(* Collect hmi signals *)
stgGr05HMI.stPLCTOHMI.bHomeCompleted := bgGr05HomeCompleted;
stgGr05HMI.stPLCTOHMI.wBtnStartStatus.0 := bgGr05StartProcess;
stgGr05HMI.stPLCTOHMI.wBtnStopStatus.0 := NOT bgGr05StartProcess;
stgGr05HMI.stPLCTOHMI.wBtnStepProcStatus := 0;
stgGr05HMI.stPLCTOHMI.wAxisClampStatus.0 := NOT binGr05AxisClamp1LimitMin;
stgGr05HMI.stPLCTOHMI.wAxisClampStatus.1 := NOT binGr05AxisClamp1LimitMax;
stgGr05HMI.stPLCTOHMI.wSlideStatus.0 := binGr05SlideTop;
stgGr05HMI.stPLCTOHMI.wSlideStatus.1 := binGr05SlideBottom;
stgGr05HMI.stPLCTOHMI.wRemovalBandStatus.0 := NOT binGr05RemovalBandInMinus;
stgGr05HMI.stPLCTOHMI.wRemovalBandStatus.1 := NOT binGr05RemovalBandInPlus;
stgGr05HMI.stPLCTOHMI.arwClampStatus[1].0 := arbinGr05ClampOpened[1];
stgGr05HMI.stPLCTOHMI.arwClampStatus[1].1 := arbinGr05ClampClosed[1];
stgGr05HMI.stPLCTOHMI.arwClampStatus[2].0 := arbinGr05ClampOpened[2];
stgGr05HMI.stPLCTOHMI.arwClampStatus[2].1 := arbinGr05ClampClosed[2];
stgGr05HMI.stPLCTOHMI.arwCylinderPosStatus[1].0 := arbinGr05CylinderPosOpened[1];
stgGr05HMI.stPLCTOHMI.arwCylinderPosStatus[1].1 := arbinGr05CylinderPosClosed[1];
stgGr05HMI.stPLCTOHMI.arwCylinderPosStatus[2].0 := arbinGr05CylinderPosOpened[2];
stgGr05HMI.stPLCTOHMI.arwCylinderPosStatus[2].1 := arbinGr05CylinderPosClosed[2];
stgGr05HMI.stPLCTOHMI.arwCylinderPosStatus[3].0 := arbinGr05CylinderPosOpened[3];
stgGr05HMI.stPLCTOHMI.arwCylinderPosStatus[3].1 := arbinGr05CylinderPosClosed[3];
stgGr05HMI.stPLCTOHMI.unSawingStep := Gr05Auto.fbProcedure.unProcessCounter;
END_ACTION

END_PROGRAM

// ---- POUs/Tc2 Objects/MachineEquipment/F_AxisClamp2Pos.TcPOU
FUNCTION F_AxisClamp2Pos : LREAL
(*

The function  used to generate position position dependent of diameter and angle.

Constructor: 		Patryk Panylo
Company:		E. Riexinger GmbH
Date:			01.04.2015
Version:			1.00

Date:			Revision:		Who:				Comment
dd.mm.yyyy		x.xx			Initials			comment

*)
VAR_INPUT
	(* Input variables / Eingang Variablen *)
	bEnable							:BOOL;						(* Function block enable *)
	lrActClamp2Pos					:LREAL;
	lrAngle							:LREAL;
	lrRadius							:LREAL;
	lrPipeClampWidth					:LREAL;
	lrSawbandGuideWidth				:LREAL;
END_VAR
VAR
	lrOffset : LREAL;
END_VAR

IF NOT bEnable
THEN
	F_AxisClamp2Pos := lrActClamp2Pos;
	RETURN;
END_IF

lrAngle := LIMIT(-45, lrAngle, 45);



F_AxisClamp2Pos := (TAN(ABS(lrAngle)) * (lrRadius + lrPipeClampWidth))
				     + (lrSawbandGuideWidth / 2 / COS(ABS(lrAngle)))
				     - (lrSawbandGuideWidth / 2);

END_FUNCTION

// ---- POUs/Tc2 Objects/Basics/FB_CheckArrayBounds.TcPOU
FUNCTION_BLOCK FB_CheckArrayBounds
VAR_INPUT
	diArrayIndex: DINT;
	diLowerBound: DINT;
	diUpperBound: DINT;
END_VAR
VAR_OUTPUT
	sLogMessage: STRING;
	diReturnBound: DINT;
END_VAR
VAR
	bErrorUpper: BOOL;
	bErrorLower: BOOL;
	fbRTrig_MessageOutputLower: R_TRIG;
	fbRTrig_MessageOutputUpper: R_TRIG;
END_VAR

(*++++++++++ Checkbounds ++++++++++*)
(*If somehow it happens that a value of any of the used arrays that does not exist is being accessed,
the value is either set to the highest declared value (if a value higher than the highest declared value is being accessed) 
or it is set to the lowest declared value (if a value lower than the lowest declared value is being accessed)  *)

IF diArrayIndex< diLowerBound THEN
	diReturnBound:= diLowerBound;
	bErrorLower:= TRUE;

	sLogMessage:= 'CheckBounds: Array index too LOW! Lower Bound: ';			(*Message is put together*)
	sLogMessage:=CONCAT(sLogMessage,DINT_TO_STRING(diLowerBound));
	sLogMessage:=CONCAT(sLogMessage,' Index being accessed: ');
	sLogMessage:=CONCAT(sLogMessage,DINT_TO_STRING(diArrayIndex));

ELSIF diArrayIndex> diUpperBound THEN
	diReturnBound:= diUpperBound;
	bErrorUpper:= TRUE;

	sLogMessage:= 'CheckBounds: Array index too HIGH! Upper Bound: ';			(*Message is put together*)
	sLogMessage:=CONCAT(sLogMessage,DINT_TO_STRING(diUpperBound));
	sLogMessage:=CONCAT(sLogMessage,' Index being accessed: ');
	sLogMessage:=CONCAT(sLogMessage,DINT_TO_STRING(diArrayIndex));

ELSIF NOT (diArrayIndex< diLowerBound) AND
	NOT (diArrayIndex> diUpperBound) THEN
		diReturnBound:= diArrayIndex;
		bErrorUpper:= FALSE;
		bErrorLower:= FALSE;
END_IF

(*++++++++++ ADSLOGDINT ++++++++++*)
(*If somehow it happens that a value of any of the used arrays that does not exist is being accessed,
the Error is written into the Logger Box of the TC System Manager  *)

fbRTrig_MessageOutputLower( CLK:= bErrorLower, Q=> );
fbRTrig_MessageOutputUpper( CLK:= bErrorUpper, Q=> );

IF fbRTrig_MessageOutputLower.Q OR fbRTrig_MessageOutputUpper.Q THEN
	ADSLOGDINT( ADSLOG_MSGTYPE_ERROR OR ADSLOG_MSGTYPE_LOG,sLogMessage,0);	(*Message is written into Event Log*)
END_IF

END_FUNCTION_BLOCK

// ---- POUs/Tc2 Objects/Basics/CheckBounds.TcPOU
FUNCTION CheckBounds : DINT
VAR_INPUT
	index: DINT;
	lower: DINT;
	upper: DINT;
END_VAR
VAR_EXTERNAL
	fbCheckArrayBounds: FB_CheckArrayBounds;
END_VAR

(*This function checks if an index out of range an array is being accessed *)

fbCheckArrayBounds(
	diArrayIndex			:= index,
	diLowerBound		:= lower,
	diUpperBound		:= upper,
	sLogMessage		=> ,
	diReturnBound		=> CheckBounds);

END_FUNCTION

// ---- POUs/Tc2 Objects/Basics/FB_CheckDivRealInfo.TcPOU
FUNCTION_BLOCK FB_CheckDivRealInfo
VAR_INPUT
	rDivisor: REAL;
END_VAR
VAR_OUTPUT
	rReturnDivReal: REAL;
	sLogMessage: STRING;
END_VAR
VAR
	bDivisorError: BOOL;
	fbRTrig_MessageOutputDiv: R_TRIG;
END_VAR

IF rDivisor= 0 THEN
	bDivisorError:= TRUE;
	rReturnDivReal:= 1;
ELSE
	rReturnDivReal:= rDivisor;
	bDivisorError:= FALSE;
END_IF

(*++++++++++ ADSLOGDINT ++++++++++*)
(*If somewhere a division by 0 is performed, an Error is written into the Logger Box of the TC System Manager  *)

fbRTrig_MessageOutputDiv( CLK:= bDivisorError, Q=> );

IF fbRTrig_MessageOutputDiv.Q THEN
	sLogMessage:= 'CheckDivReal Error: Division by Zero! Divisor set from 0 to 1. ';					(*Message*)

	ADSLOGDINT( ADSLOG_MSGTYPE_ERROR OR ADSLOG_MSGTYPE_LOG,sLogMessage,0);	(*Message is written into Event Log*)
END_IF

END_FUNCTION_BLOCK

// ---- POUs/Tc2 Objects/Basics/CheckDivReal.TcPOU
FUNCTION CheckDivReal : REAL
VAR_INPUT
	divisor: REAL;
END_VAR
VAR_EXTERNAL
	fbCheckDivRealInfo: FB_CheckDivRealInfo;
END_VAR

(*This function checks if a division by zero is performed*)

fbCheckDivRealInfo(
	rDivisor			:= divisor,
	sLogMessage	=> ,
	rReturnDivReal 	=> CheckDivReal);

END_FUNCTION

// ---- POUs/FAST.TcPOU
PROGRAM FAST
VAR
	(* Enummerations *)

	(* Variables *)

	(* References *)

	(* Interfaces *)

	(* Instances *)

END_VAR


;

END_PROGRAM

// ---- POUs/Tc2 Objects/Automation/Axis/Beckhoff/FB_AxisMcBeckhoff.TcPOU
FUNCTION_BLOCK FB_AxisMcBeckhoff
(*

The function block used to control axis welding.

Constructor: 		Patryk Panylo
Company:		E. Riexinger GmbH
Date:			28.04.2015
Version:			1.00

Date:			Revision:		Who:				Comment
dd.mm.yyyy		x.xx			Initials			comment

*)
VAR_INPUT
	(* Input variables / Eingang Variablen *)
	bEnable						:BOOL;						(* Axis present *)
	etMachineMode				:ET_MachineMode;			(* Machine mode *)
	etMachineState				:ET_MachineState;			(* Machine state *)
	bNoEStop					:BOOL;						(* No ermergency Stop / Keine Notaus *)
	bPowerSupplyOn				:BOOL;						(* Power supply on / Leitung eingeschaltet *)
	bLightCurtainOK				:BOOL;						(* Light curtain ok / Freigabe Lichtschranke i.o *)
	bMachineStandstill			:BOOL;						(* Machine standstill *)
	bCtrlInterrupt					:BOOL;						(* Control interrupt *)
	bMoveRelease				:BOOL;						(* Move release *)
	lrSoftLimitMax					:LREAL; 						(* Position limit switch maximum *)
	lrSoftLimitMin					:LREAL; 						(* Position limit switch minimum *)
	bTipPlus						:BOOL;						(* Manual tip in plus direction *)
	bTipMinus					:BOOL;						(* Manual tip in minus direction *)
	lrTipDistance					:LREAL;						(* Relative distance for movements *)
	bPlusRelease				:BOOL;						(* Plus move release *)
	bMinusRelease				:BOOL;						(* Minus move release *)
	bExeSetPos					:BOOL;						(* Execute set position *)
	bExeHome					:BOOL;						(* Execute home *)
	etHomingMode 				:MC_HomingMode;			(* HomingMode determines in which way the calibration is carried out. *)
	bExeMoveAbs				:BOOL;						(* Execute move absolut *)
	bExeMoveRel				:BOOL;						(* Execute move relative *)
	bExeMoveAdd				:BOOL;						(* Execute move additive *)
	bExeMoveSuper				:BOOL;						(* Execute move superimposed *)
	bExeMoveVelo				:BOOL;						(* Execute move velo *)
	bExeGearIn					:BOOL;						(* Execute gear in *)
	bExeGearOut					:BOOL;						(* Execute gear out *)
	bExeStop					:BOOL;						(* Execute move stop *)
	bExeReset					:BOOL;						(* Execute auto reset *)
	bExtOverrideEn				:BOOL;						(* External override enable *)
	lrExtOverride					:LREAL;						(* External override *)
	lrTargetPosition				:LREAL;						(* Absolute target position *)
	lrManualVelocity				:LREAL;						(* Value of velocity in manual motion [mm/s] *)
	lrVelocityNoRef				:LREAL;						(* Velocity if has no reference [mm/s] *)
	bVelocityLimitEn				:BOOL;						(* Enable velocity limit *)
	lrAutoVelocity					:LREAL;						(* Value of velocity in auto motion [mm/s] *)
	lrVelocityMin					:LREAL;						(* Velocity minimum [%] *)
	lrVelocityMax					:LREAL;						(* Velocity maximum [%] *)
	lrAcceleration					:LREAL;						(* Value of the acceleration (always positive). If >= 0 else from SM *)
	lrDeceleration				:LREAL;						(* Value of deceleration (always positive). If >= 0 else from SM *)
	lrJerk						:LREAL;						(* Value of jerk (always positive). If >= 0 else from SM *)
	bEngineTorqueLimitEn			:BOOL;						(* Enable engine torque limit *)
	lrEngineTorque				:LREAL;						(* Engine torque [%] *)
	bWithAbsoluteEncoder			:BOOL; 						(* Encoder is an absolute one / Absolutwertgeber *)
	bPosLagMonitoringEn			:BOOL;						(* Enable position lag monitoring *)
	lrOriginShiftPos				:LREAL;						(* Origin shift position *)
	dnRatioNumerator				:DINT;						(* Gear ratio numerator. Alternatively, the gear ratio can be specified in the numerator as a floating comma value, if the denominator is 1. *)
	udnRatioDenominator			:UDINT;						(* Gear ratio denominator *)
	bVeloForceCtrlEn				:BOOL;						(* Enable velocity  force controller *)
	lrVeloForceCtrlKp				:LREAL;						(* Velocity - force controller proportional band Kp *)
	lrVeloForceCtrlTi				:LREAL;						(* Velocity - force controller integral Ti *)
	lrVeloForceCtrlMin				:LREAL;						(* Velocity - force controller minimum  *)
	lrVeloForceCtrlMax			:LREAL;						(* Velocity - force controller maxmimum  *)
	lrTargetForce					:LREAL;						(* Absolute target force [N] *)
	lrForceCurrent				:LREAL;						(* Current force [mA] *)
	rForceOffset					:REAL;						(* Force offset [N] *)
	lrForceMinmA					:LREAL;						(* Force min [mA] 16#0000 = 4 [mA] *)
	lrForceMaxmA 				:LREAL;						(* Force max [mA] 16#7FFF = 20 [mA] *)
	lrForceMinN					:LREAL;						(* Force min [N] *)
	lrForceMaxN					:LREAL;						(* Force max [N] *)
	lrOverride					:LREAL;						(* Override *)
	lrActTemp					:LREAL;						(* Current temperatur *)
	lrTempLimitMax				:LREAL;						(* Temperatur limit maximum*)
	lrTempLimitMin				:LREAL;						(* Temperatur limit minimum*)
	bCoolingActive				:BOOL;						(* Cooling on *)
	bConfirmAlarm				:BOOL;						(* Confirm alarm *)
	bOccupied					:BOOL;						(* Axis occupied *)
	tControllerOff					:TIME := t#60s;				(* Time to switch controller off *)
	tAdsTimeOut 					:TIME := t#2s;					(* Timout for ads commands *)
END_VAR
VAR_OUTPUT
	(* Output variables / Ausgang Variablen *)
	bCtrlEnabled					:BOOL;						(* Controller enabled *)
	bNotMoving					:BOOL;						(* Axis not moving *)
	bReferenced					:BOOL;						(* Axis referenced *)
	bCoupled					:BOOL;						(* Axis coupled *)
	lrActPosition					:LREAL;						(* Actual position [mm] *)
	lrActAbsPosition				:LREAL;						(* Actual absolut position [mm] *)
	lrActVelocity					:LREAL;						(* Actual velocity [mm/s] *)
	lrActForce					:LREAL;						(* Actual force [N] *)
	lrVeloMax					:LREAL;						(* Velocity limit maximum *)
	lrAccMax						:LREAL;						(* Acceleration limit maximum *)
	lrDecMax					:LREAL;						(* Deceleration limit maximum *)
	lrJerkMax					:LREAL;						(* Jerk limit maximum *)
	bHardLimitMaxExceeded		:BOOL;						(* Position limit switch maximum is exceeded *)
	bHardLimitMinExceeded		:BOOL;						(* Position limit switch minimum is exceeded *)
	bSoftLimitMaxExceeded		:BOOL;						(* Position limit switch maximum is exceeded *)
	bSoftLimitMinExceeded		:BOOL;						(* Position limit switch minimum is exceeded *)
	bCoolingOn					:BOOL;						(* Cooling *)
	bErrorTerminal				:BOOL;						(* Error Axis terminal *)
	bErrorCtrlEnabled				:BOOL;						(* Error Axis controller enabled *)
END_VAR
VAR_IN_OUT
	(* Input Output variables / Ausgang Variablen *)
	bHomeCompleted				:BOOL;						(* Home completed *)
	Drive						:ST_BECKHOFFDRIVE_REF; 	(* The ST_BECHOFFDRIVE_REF data type  is an interface between the PLC and the DRIVE and contains axis information *)
	Axis							:AXIS_REF;					(* The AXIS_REF data type  is an interface between the PLC and the NC and contains axis information *)
	MasterAxis					:AXIS_REF;					(* The AXIS_REF data type  is an interface between the PLC and the NC and contains axis information *)
END_VAR
VAR
	(* Enummerations *)

	(* Variables *)
	sAdsAddr					:STRING(23);					(* AmsNetId of the EtherCAT master device.*)
	unSlaveAddr					:UINT;						(* Address of the slave device.*)

	nTorqueLimitMax				:INT := 100;					(* The torque limit (absolute value). Value range in %: -200 ... 200 ... 200 *)

	lrVeloLimitMax				:LREAL;
	lrVeloLimitMin					:LREAL;

	sTerminalStatus				:STRING;
	(* References *)

	(* Interfaces *)

	(* Instances *)
	fbTerminalDiagnosis			:FB_TerminalDiagnosis;
	rtMachineStandstill			:R_TRIG;
	tonAxisEnabled				:TON;

	fbController					:FB_AxisController;
	fbMoveManual				:FB_AxisMoveManual;
	fbMoveAuto					:FB_AxisMoveAuto;
	fbForce						:FB_ScalingOffset;
	fbForceCtrl					:FB_ForceController;
	fbCoolingOff					:FB_SignalHandlingDelay;
END_VAR


IF NOT bEnable								(* Signal FB enable *)
THEN

	RETURN;
END_IF

A_AxisLink();
A_AxisGetStatus();
A_AxisController();
A_AxisForceCtrl();
A_AxisMoveManual();
A_AxisMoveAuto();
A_AxisCooling();
A_AxisTerminalDiag();
A_AxisAlarm();

ACTION A_AxisAlarm:

(* Axis errors *)
tonAxisEnabled(
	IN := fbController.bEnable
		AND fbController.bRegulatorOn
		AND NOT fbController.bStatusDelay,
	PT := fbController.tStatusDelay + t#2s
);

bErrorCtrlEnabled := tonAxisEnabled.Q;
END_ACTION

ACTION A_AxisController:

(* Axis controller *)
fbController(
    	bEnable := TRUE,
	etMachineMode := etMachineMode,
	etMachineState := etMachineState,
	bRegulatorOn := bNoEStop
				      AND bPowerSupplyOn
				      AND bLightCurtainOK
				      AND SEL(bNotMoving, NOT bCtrlInterrupt, TRUE)
				      AND NOT fbMoveManual.bControllerOff
				      AND NOT fbMoveAuto.bControllerOff ,
	bReset := bConfirmAlarm,
	bTerminalOK := fbTerminalDiagnosis.bTerminalOK,
	bExeReset := bExeReset,
	bExeSetPos := bExeSetPos,
	lrSetPosition := lrTargetPosition,
	bExeGearIn := bExeGearIn,
	bExeGearOut := bExeGearOut,
	dnRatioNumerator := dnRatioNumerator,
	udnRatioDenominator := udnRatioDenominator,
	lrOverride := SEL(bExtOverrideEn,
					SEL(
						bVeloForceCtrlEn,
						lrOverride,
						fbForceCtrl.lrCVVelo),
					lrOverride*lrExtOverride/100.0),
	bWithAbsoluteEncoder := bWithAbsoluteEncoder,
	bPosLagMonitoringEn := bPosLagMonitoringEn,
	lrPositionBias := lrOriginShiftPos,
	lrSoftLimitMax := lrSoftLimitMax,
	lrSoftLimitMin := lrSoftLimitMin,
	lrAcceleration := lrAcceleration,
	lrDeceleration := lrDeceleration,
	lrJerk := lrJerk,
	Axis := Axis,
	MasterAxis := MasterAxis,
	bStatusDelay => bCtrlEnabled,
	lrActPos => lrActPosition,
	lrActAbsPos => lrActAbsPosition,
	lrActVelo => lrActVelocity,
	bNotMoving => bNotMoving,
	bReferenced => bReferenced,
	bCoupled => bCoupled,
	lrVeloLimitMax => lrVeloMax,
	lrAccLimitMax => lrAccMax,
	lrDecLimitMax => lrDecMax,
	lrJerkLimitMax => lrJerkMax,
	bHardLimitMaxExceeded => bHardLimitMaxExceeded,
	bHardLimitMinExceeded => bHardLimitMinExceeded,
	bSoftLimitMaxExceeded => bSoftLimitMaxExceeded,
	bSoftLimitMinExceeded => bSoftLimitMinExceeded
);
END_ACTION

ACTION A_AxisCooling:

(* Cooling control *)
fbCoolingOff(
	bEnable := TRUE,
	bIn := NOT bCoolingActive
		  AND lrActTemp < lrTempLimitMin
		  AND bCoolingOn,
	tDelay := t#30s
);

IF bCoolingActive
     OR lrActTemp > lrTempLimitMax
THEN
	bCoolingOn := TRUE;

ELSIF fbCoolingOff.bOut
THEN
	bCoolingOn := FALSE;
END_IF
END_ACTION

ACTION A_AxisForceCtrl:

fbForce(
	bEnable := TRUE,
	lrInput := lrForceCurrent,
	lrXLowLimit := lrForceMinmA, (* 16#0000 = 4 [mA] *)
	lrXUpperLimit := lrForceMaxmA, (* 16#7FFF = 20 [mA] *)
	lrYLowLimit := lrForceMinN,  (*[N]*)
	lrYUpperLimit := lrForceMaxN,  (*[N]*)
	usiPrecision := 2,
	lrOffset := rForceOffset,
	lrOutputPV => lrActForce
);

fbForceCtrl(
	bEnable := bNoEStop
			    AND bPowerSupplyOn
			    AND bLightCurtainOK
			    AND bCtrlEnabled,
	bControllerOn := bVeloForceCtrlEn,
	lrVeloKp := lrVeloForceCtrlKp,
	lrVeloTi := lrVeloForceCtrlTi,
	lrPVForce := lrActForce, (* [N] *)
	lrSPForce := lrTargetForce, (* [N] *)
	lrMaxForce := lrForceMaxN, (* [N] *)
	lrVeloMax := lrVeloForceCtrlMax,
	lrVeloMin := lrVeloForceCtrlMin,
	lrTaskCycle := lrgActCycleTime
);
END_ACTION

ACTION A_AxisGetStatus:

(* Get axis status *)
Axis.ReadStatus();
END_ACTION

ACTION A_AxisLink:

(* Get terminal status *)
sAdsAddr:= F_CreateAmsNetId(Drive.stTerminalState.stAdsAddr.netId);
unSlaveAddr:= Drive.stTerminalState.stAdsAddr.port;

(* Set drive parameter *)
(*Drive.stPlcToStoeber.snA541ModesOfOperation := snModesOfOperation;*)

(*Drive.PlcToStoeber.nA558TargetTorque := SEL(bEngineTorqueLimitEn,
				    nTorqueLimitMax,
				    LREAL_TO_INT(lrEngineTorque / 1.0))*)
END_ACTION

ACTION A_AxisMoveAuto:

(* Move axis auto *)
rtMachineStandstill(CLK := bMachineStandstill );

lrVeloLimitMin := SEL(bVelocityLimitEn, -1 * lrVeloMax, lrVelocityMin);
lrVeloLimitMax := SEL(bVelocityLimitEn, lrVeloMax, lrVelocityMax);

fbMoveAuto(
	bEnable := bNoEStop
               		    AND bPowerSupplyOn
               		    AND bLightCurtainOK,
	bOccupied := bOccupied,
	bCtrlEnabled := bCtrlEnabled
				      AND bMoveRelease,
	etMachineMode := etMachineMode,
	etMachineState := etMachineState,
	bReset := bConfirmAlarm,
	bExeHome := bExeHome,
	bExeMoveAbs := bExeMoveAbs,
	bExeMoveRel := bExeMoveRel,
	bExeMoveAdd := bExeMoveAdd,
	bExeMoveSuper := bExeMoveSuper,
	bExeMoveVelo := bExeMoveVelo,
	bExeStop := bExeStop
			      OR rtMachineStandstill.Q,
	etHomingMode := etHomingMode,
	lrPosition := lrTargetPosition,
	lrVelocity := LIMIT(lrVeloLimitMin, lrAutoVelocity, lrVeloLimitMax),
	lrAcceleration := lrAcceleration,
	lrDeceleration := lrDeceleration,
	lrJerk := lrJerk,
	lrOriginShiftPos := lrOriginShiftPos,
	bSignalReference := (*Drive.stStoeberToPlc.dw1A636DigitalInputs.2*),
	tControllerOff := tControllerOff,
	bHomeCompleted := bHomeCompleted,
	Axis := Axis,
	MasterAxis := MasterAxis
 );
END_ACTION

ACTION A_AxisMoveManual:

(* Move axis manual *)
fbMoveManual(
	bEnable := bNoEStop
               		    AND bPowerSupplyOn
               		    AND bLightCurtainOK,
	bOccupied := bOccupied,
	bCtrlEnabled := bCtrlEnabled
				      AND bMoveRelease,
	etMachineMode := etMachineMode,
	etMachineState := etMachineState,
	bReset := bConfirmAlarm,
	bMovePlus := bTipPlus,
	bMoveMinus := bTipMinus,
	lrTipDistance := lrTipDistance,
	bLimitMax := bHardLimitMaxExceeded
			       OR bSoftLimitMaxExceeded,
	bLimitMin := bHardLimitMinExceeded
			      OR bSoftLimitMinExceeded,
	bPlusRelease := bPlusRelease,
	bMinusRelease := bMinusRelease,
	lrVelocity := SEL(NOT bReferenced, lrManualVelocity, lrVelocityNoRef),
	lrAcceleration := lrAcceleration,
	lrDeceleration := lrDeceleration,
	lrJerk := lrJerk,
	tControllerOff := tControllerOff,
	bHomeCompleted := bHomeCompleted,
	Axis := Axis,
	MasterAxis := MasterAxis
);
END_ACTION

ACTION A_AxisTerminalDiag:

(*Axis terminal diagnosis *)
fbTerminalDiagnosis(
	stTerminalState := Drive.stTerminalState,
	sTerminalStatus => sTerminalStatus
);

bErrorTerminal := NOT fbTerminalDiagnosis.bTerminalOK;
END_ACTION

END_FUNCTION_BLOCK

// ---- POUs/Tc2 Objects/Automation/Axis/Beckhoff/FB_AxisMcBeckhoffSEWMoviDriveBVelo.TcPOU
FUNCTION_BLOCK FB_AxisMcBeckhoffSEWMoviDriveBVelo
(*

The function block used to control axis welding.

Constructor: 		Patryk Panylo
Company:		E. Riexinger GmbH
Date:			28.04.2015
Version:			1.00

Date:			Revision:		Who:				Comment
dd.mm.yyyy		x.xx			Initials			comment

*)
VAR_INPUT
	(* Input variables / Eingang Variablen *)
	bEnable						:BOOL;						(* Axis present *)
	etMachineMode				:ET_MachineMode;			(* Machine mode *)
	etMachineState				:ET_MachineState;			(* Machine state *)
	bNoEStop					:BOOL;						(* No ermergency Stop / Keine Notaus *)
	bPowerSupplyOn				:BOOL;						(* Power supply on / Leitung eingeschaltet *)
	bLightCurtainOK				:BOOL;						(* Light curtain ok / Freigabe Lichtschranke i.o *)
	bMachineStandstill			:BOOL;						(* Machine standstill *)
	bCtrlInterrupt					:BOOL;						(* Control interrupt *)
	bMoveRelease				:BOOL;						(* Move release *)
	lrSoftLimitMax					:LREAL; 						(* Position limit switch maximum *)
	lrSoftLimitMin					:LREAL; 						(* Position limit switch minimum *)
	bTipPlus						:BOOL;						(* Manual tip in plus direction *)
	bTipMinus					:BOOL;						(* Manual tip in minus direction *)
	lrTipDistance					:LREAL;						(* Relative distance for movements *)
	bPlusRelease				:BOOL;						(* Plus move release *)
	bMinusRelease				:BOOL;						(* Minus move release *)
	bExeSetPos					:BOOL;						(* Execute set position *)
	bExeHome					:BOOL;						(* Execute home *)
	etHomingMode 				:MC_HomingMode;			(* HomingMode determines in which way the calibration is carried out. *)
	bExeMoveAbs				:BOOL;						(* Execute move absolut *)
	bExeMoveRel				:BOOL;						(* Execute move relative *)
	bExeMoveAdd				:BOOL;						(* Execute move additive *)
	bExeMoveSuper				:BOOL;						(* Execute move superimposed *)
	bExeMoveVelo				:BOOL;						(* Execute move velo *)
	bExeGearIn					:BOOL;						(* Execute gear in *)
	bExeGearOut					:BOOL;						(* Execute gear out *)
	bExeStop					:BOOL;						(* Execute move stop *)
	bExeReset					:BOOL;						(* Execute auto reset *)
	bExtOverrideEn				:BOOL;						(* External override enable *)
	lrExtOverride					:LREAL;						(* External override *)
	lrTargetPosition				:LREAL;						(* Absolute target position *)
	lrManualVelocity				:LREAL;						(* Value of velocity in manual motion [mm/s] *)
	lrVelocityNoRef				:LREAL;						(* Velocity if has no reference [mm/s] *)
	bVelocityLimitEn				:BOOL;						(* Enable velocity limit *)
	lrAutoVelocity					:LREAL;						(* Value of velocity in auto motion [mm/s] *)
	lrVelocityMin					:LREAL;						(* Velocity minimum [%] *)
	lrVelocityMax					:LREAL;						(* Velocity maximum [%] *)
	lrAcceleration					:LREAL;						(* Value of the acceleration (always positive). If >= 0 else from SM *)
	lrDeceleration				:LREAL;						(* Value of deceleration (always positive). If >= 0 else from SM *)
	lrJerk						:LREAL;						(* Value of jerk (always positive). If >= 0 else from SM *)
	bEngineTorqueLimitEn			:BOOL;						(* Enable engine torque limit *)
	lrEngineTorque				:LREAL;						(* Engine torque [%] *)
	bWithAbsoluteEncoder			:BOOL; 						(* Encoder is an absolute one / Absolutwertgeber *)
	bPosLagMonitoringEn			:BOOL;						(* Enable position lag monitoring *)
	lrOriginShiftPos				:LREAL;						(* Origin shift position *)
	dnRatioNumerator				:DINT;						(* Gear ratio numerator. Alternatively, the gear ratio can be specified in the numerator as a floating comma value, if the denominator is 1. *)
	udnRatioDenominator			:UDINT;						(* Gear ratio denominator *)
	bVeloForceCtrlEn				:BOOL;						(* Enable velocity - force controller *)
	lrVeloForceCtrlKp				:LREAL;						(* Velocity - force controller proportional band Kp *)
	lrVeloForceCtrlTi				:LREAL;						(* Velocity - force controller integral Ti *)
	lrVeloForceCtrlVeloFilter		:LREAL;						(* Velocity control filter wieghting =  0..1 *)
	lrVeloForceCtrlLimit			:LREAL;						(* Velocity - force controller limit  *)
	lrTargetForce					:LREAL;						(* Absolute target force [N] *)
	lrForceCurrent				:LREAL;						(* Current force [mA] *)
	lrForceOffset					:LREAL;						(* Force offset [N] *)
	lrOverride					:LREAL;						(* Override *)
	lrActTemp					:LREAL;						(* Current temperatur *)
	lrTempLimitMax				:LREAL;						(* Temperatur limit maximum*)
	lrTempLimitMin				:LREAL;						(* Temperatur limit minimum*)
	bCoolingActive				:BOOL;						(* Cooling on *)
	bConfirmAlarm				:BOOL;						(* Confirm alarm *)
	bOccupied					:BOOL;						(* Axis occupied *)
	tControllerOff					:TIME := t#60s;				(* Time to switch controller off *)
	tAdsTimeOut 					:TIME := t#2s;					(* Timout for ads commands *)
END_VAR
VAR_OUTPUT
	(* Output variables / Ausgang Variablen *)
	bCtrlEnabled					:BOOL;						(* Controller enabled *)
	bNotMoving					:BOOL;						(* Axis not moving *)
	bReferenced					:BOOL;						(* Axis referenced *)
	bCoupled					:BOOL;						(* Axis coupled *)
	lrActPosition					:LREAL;						(* Actual position [mm] *)
	lrActAbsPosition				:LREAL;						(* Actual absolut position [mm] *)
	lrActVelocity					:LREAL;						(* Actual velocity [mm/s] *)
	lrActForce					:LREAL;						(* Actual force [N] *)
	lrVeloMax					:LREAL;						(* Velocity limit maximum *)
	lrAccMax						:LREAL;						(* Acceleration limit maximum *)
	lrDecMax					:LREAL;						(* Deceleration limit maximum *)
	lrJerkMax					:LREAL;						(* Jerk limit maximum *)
	bHardLimitMaxExceeded		:BOOL;						(* Position limit switch maximum is exceeded *)
	bHardLimitMinExceeded		:BOOL;						(* Position limit switch minimum is exceeded *)
	bSoftLimitMaxExceeded		:BOOL;						(* Position limit switch maximum is exceeded *)
	bSoftLimitMinExceeded		:BOOL;						(* Position limit switch minimum is exceeded *)
	bCoolingOn					:BOOL;						(* Cooling *)
	bErrorTerminal				:BOOL;						(* Error Axis terminal *)
	bErrorDrive					:BOOL;						(* Error drive *)
	bErrorCtrlEnabled				:BOOL;						(* Error Axis controller enabled *)
	bErrorForce					:BOOL;						(* Error force *)
END_VAR
VAR_IN_OUT
	(* Input Output variables / Ausgang Variablen *)
	bHomeCompleted				:BOOL;						(* Home completed *)
	Drive						:ST_SEWMOVIEDRIVEBCIA402_REF; (* The ST_SEWMOVIEDRIVEBCIA402_REF data type  is an interface between the PLC and the DRIVE and contains axis information *)
	Axis							:AXIS_REF;					(* The AXIS_REF data type  is an interface between the PLC and the NC and contains axis information *)
	MasterAxis					:AXIS_REF;					(* The AXIS_REF data type  is an interface between the PLC and the NC and contains axis information *)
	Force						:ST_FORCE_REF; 			(* The ST_FORCE_REF data type  is an interface between the PLC and the FORCE and contains axis information *)
END_VAR
VAR
	(* Enummerations *)

	(* Variables *)
	sAdsAddr					:STRING(23);					(* AmsNetId of the EtherCAT master device.*)
	unSlaveAddr					:UINT;						(* Address of the slave device.*)

	nTorqueLimitMax				:INT := 100;					(* The torque limit (absolute value). Value range in %: -200 ... 200 ... 200 *)

	lrVeloLimitMax				:LREAL;
	lrVeloLimitMin					:LREAL;

	sTerminalStatus				:STRING;

	bSetDefaultSettings			:BOOL;
	bReadSettings				:BOOL;
	bWriteSettings				:BOOL;

	rCacheWeightTara			:REAL;

	(* References *)

	(* Interfaces *)

	(* Instances *)
	fbTerminalDiagnosis			:FB_TerminalDiagnosis;
	rtMachineStandstill			:R_TRIG;
	tonAxisEnabled				:TON;

	fbController					:FB_AxisController;
	fbMoveManual				:FB_AxisMoveManual;
	fbMoveAuto					:FB_AxisMoveAuto;
	fbForceCtrl					:FB_ForceController;
	fbCoolingOff					:FB_SignalHandlingDelay;
END_VAR


IF NOT bEnable								(* Signal FB enable *)
THEN

	RETURN;
END_IF

A_AxisLink();
A_AxisGetStatus();
A_AxisController();
A_AxisForceCtrl();
A_AxisMoveManual();
A_AxisMoveAuto();
A_AxisCooling();
A_AxisTerminalDiag();
A_AxisAlarm();

ACTION A_AxisAlarm:

(* Axis errors *)
tonAxisEnabled(
	IN := fbController.bEnable
		AND fbController.bRegulatorOn
		AND NOT fbController.bStatusDelay,
	PT := fbController.tStatusDelay + t#2s
);

bErrorCtrlEnabled := tonAxisEnabled.Q;

bErrorForce := ((etMachineMode = ET_MachineMode_eAutomatic
			    OR etMachineMode = ET_MachineMode_eHome) AND lrActForce > Force.lrAutoForceMaxN)
			  OR (etMachineMode = ET_MachineMode_eManual AND lrActForce > Force.lrManualForceMaxN);
END_ACTION

ACTION A_AxisController:

(* Axis controller *)
fbController(
    	bEnable := TRUE,
	etMachineMode := etMachineMode,
	etMachineState := etMachineState,
	bRegulatorOn := bNoEStop
				      AND bPowerSupplyOn
				      AND bLightCurtainOK
				      AND SEL(bNotMoving, NOT bCtrlInterrupt, TRUE)
				      AND Drive.stSEWToPlc.wPO1StatusWord.1			(* Umrichter betriebsbereit *)
				      AND Drive.stSEWToPlc.wPO1StatusWord.2			(* PA-Daten freigegeben *)
				      AND NOT fbMoveManual.bControllerOff
				      AND NOT fbMoveAuto.bControllerOff ,
	bReset := bConfirmAlarm,
	bTerminalOK := fbTerminalDiagnosis.bTerminalOK,
	bExeReset := bExeReset,
	bExeSetPos := bExeSetPos,
	lrSetPosition := lrTargetPosition,
	bExeGearIn := bExeGearIn,
	bExeGearOut := bExeGearOut,
	dnRatioNumerator := dnRatioNumerator,
	udnRatioDenominator := udnRatioDenominator,
	lrOverride := SEL(bExtOverrideEn,
					SEL(
						bVeloForceCtrlEn,
						lrOverride,
						fbForceCtrl.lrCVVelo),
					lrOverride*lrExtOverride/100.0),
	bWithAbsoluteEncoder := bWithAbsoluteEncoder,
	bPosLagMonitoringEn := bPosLagMonitoringEn,
	lrPositionBias := lrOriginShiftPos,
	bHWSignalLimitMax := NOT Drive.stSEWToPlc.bAxisWeldingLimitMax,
	bHWSignalLimitMin := NOT Drive.stSEWToPlc.bAxisWeldingLimitMin,
	lrSoftLimitMax := lrSoftLimitMax,
	lrSoftLimitMin := lrSoftLimitMin,
	lrAcceleration := lrAcceleration,
	lrDeceleration := lrDeceleration,
	lrJerk := lrJerk,
	Axis := Axis,
	MasterAxis := MasterAxis,
	bStatusDelay => bCtrlEnabled,
	lrActPos => lrActPosition,
	lrActAbsPos => lrActAbsPosition,
	lrActVelo => lrActVelocity,
	bNotMoving => bNotMoving,
	bReferenced => bReferenced,
	bCoupled => bCoupled,
	lrVeloLimitMax => lrVeloMax,
	lrAccLimitMax => lrAccMax,
	lrDecLimitMax => lrDecMax,
	lrJerkLimitMax => lrJerkMax,
	bHardLimitMaxExceeded => bHardLimitMaxExceeded,
	bHardLimitMinExceeded => bHardLimitMinExceeded,
	bSoftLimitMaxExceeded => bSoftLimitMaxExceeded,
	bSoftLimitMinExceeded => bSoftLimitMinExceeded
);
END_ACTION

ACTION A_AxisCooling:

(* Cooling control *)
fbCoolingOff(
	bEnable := TRUE,
	bIn := NOT bCoolingActive
		  AND lrActTemp < lrTempLimitMin
		  AND bCoolingOn,
	tDelay := t#30s
);

IF bCoolingActive
     OR lrActTemp > lrTempLimitMax
THEN
	bCoolingOn := TRUE;

ELSIF fbCoolingOff.bOut
THEN
	bCoolingOn := FALSE;
END_IF
END_ACTION

ACTION A_AxisForceCtrl:

IF Force.unForceMeasureType = 1			(* Current or voltage force measure *)
THEN
	Force.fbForceSimple(
		bEnable := TRUE,
		lrInput := lrForceCurrent,
		lrXLowLimit := Force.lrForceMin, (* 16#0000 = 4 [mA] *)
		lrXUpperLimit := Force.lrForceMax, (* 16#7FFF = 20 [mA] *)
		lrYLowLimit := Force.lrForceMinN,  (*[N]*)
		lrYUpperLimit := Force.lrAutoForceMaxN,  (*[N]*)
		usiPrecision := 2,
		lrOffset := lrForceOffset,
		lrOutputPV => lrActForce
	);


ELSIF Force.unForceMeasureType = 2			(* EL3351 force measure *)
THEN
	;

ELSIF  Force.unForceMeasureType = 3			(* EL3356 force measure *)
THEN

	bWriteSettings := rCacheWeightTara <> Force.stRefSettingsEL3356.rTara;

	Force.fbForceEL3356(
		bEnable := TRUE,
		nTerminalNr := 1,
		stTerminalState := Force.stTerminalStateEL3356,
		stChannelState := Force.stChannelStateEL3356,
		bSetCoeParaToDefault := bSetDefaultSettings,
		bReadCoePara := bReadSettings,
		bWriteCoePara := bWriteSettings,
		rValue := lrForceCurrent,
		stCoeWrite := Force.stRefSettingsEL3356,
		stCoeRead => Force.stActSettingsEL3356,
		stChannelCtrl => Force.stChannelCtrlEL3356,
		lrGrossWeightPV =>
	);

	lrActForce := F_LRealRound(Force.fbForceEL3356.lrGrossWeightPV - lrForceOffset, 2);

	rCacheWeightTara := Force.stRefSettingsEL3356.rTara;

ELSE							(* Directly force measure *)

	lrActForce := lrForceCurrent;

END_IF

fbForceCtrl(
	bEnable := bNoEStop
			    AND bPowerSupplyOn
			    AND bLightCurtainOK
			    AND bCtrlEnabled,
	bControllerOn := bVeloForceCtrlEn,
	lrVeloKp := lrVeloForceCtrlKp,
	lrVeloTi := lrVeloForceCtrlTi,
	lrCtrlVeloFilter := lrVeloForceCtrlVeloFilter,
	lrPVForce := lrActForce, (* [N] *)
	lrSPForce := lrTargetForce, (* [N] *)
	lrMaxForce := Force.lrAutoForceMaxN, (* [N] *)
	lrVeloMax := lrVeloForceCtrlLimit,
	lrVeloMin := -lrVeloForceCtrlLimit,
	lrTaskCycle := lrgActCycleTime
);
END_ACTION

ACTION A_AxisGetStatus:

(* Get axis status *)
Axis.ReadStatus();
END_ACTION

ACTION A_AxisLink:

(* Get terminal status *)
sAdsAddr:= F_CreateAmsNetId(Drive.stTerminalState.stAdsAddr.netId);
unSlaveAddr:= Drive.stTerminalState.stAdsAddr.port;

bErrorDrive := Drive.stSEWToPlc.wPO1StatusWord.5;			(* Störung / Warnung *)

(* Set drive parameter *)
Drive.stPlcToSEW.wPO1ControlWord.1 := bCtrlEnabled;			(* Freigabe 1 / Schnellstop 0 *)
Drive.stPlcToSEW.wPO1ControlWord.2 := bCtrlEnabled;			(* Freigabe 1 / Halt 0 *)
Drive.stPlcToSEW.wPO1ControlWord.6 := bConfirmAlarm;		(* Reset *)
END_ACTION

ACTION A_AxisMoveAuto:

(* Move axis auto *)
rtMachineStandstill(CLK := bMachineStandstill);

lrVeloLimitMin := SEL(bVelocityLimitEn, -1 * lrVeloMax, lrVelocityMin);
lrVeloLimitMax := SEL(bVelocityLimitEn, lrVeloMax, lrVelocityMax);

fbMoveAuto(
	bEnable := bNoEStop
               		    AND bPowerSupplyOn
               		    AND bLightCurtainOK,
	bOccupied := bOccupied,
	bCtrlEnabled := bCtrlEnabled
				      AND bMoveRelease
				      AND Drive.stSEWToPlc.wPO1StatusWord.0,			(* Endstufe freigegeben *)
	etMachineMode := etMachineMode,
	etMachineState := etMachineState,
	bReset := bConfirmAlarm,
	bExeHome := bExeHome,
	bExeMoveAbs := bExeMoveAbs,
	bExeMoveRel := bExeMoveRel,
	bExeMoveAdd := bExeMoveAdd,
	bExeMoveSuper := bExeMoveSuper,
	bExeMoveVelo := bExeMoveVelo,
	bExeStop := bExeStop
			      OR rtMachineStandstill.Q,
	etHomingMode := etHomingMode,
	lrPosition := lrTargetPosition,
	lrVelocity := LIMIT(lrVeloLimitMin, lrAutoVelocity, lrVeloLimitMax),
	lrAcceleration := lrAcceleration,
	lrDeceleration := lrDeceleration,
	lrJerk := lrJerk,
	lrOriginShiftPos := lrOriginShiftPos,
	bSignalReference := NOT Drive.stSEWToPlc.bAxisWeldingLimitMax,
	tControllerOff := tControllerOff,
	bHomeCompleted := bHomeCompleted,
	Axis := Axis,
	MasterAxis := MasterAxis
 );
END_ACTION

ACTION A_AxisMoveManual:

(* Move axis manual *)
fbMoveManual(
	bEnable := bNoEStop
               		    AND bPowerSupplyOn
               		    AND bLightCurtainOK,
	bOccupied := bOccupied,
	bCtrlEnabled := bCtrlEnabled
				      AND bMoveRelease
				      AND Drive.stSEWToPlc.wPO1StatusWord.0,			(* Endstufe freigegeben *)
	etMachineMode := etMachineMode,
	etMachineState := etMachineState,
	bReset := bConfirmAlarm,
	bMovePlus := bTipPlus,
	bMoveMinus := bTipMinus,
	lrTipDistance := lrTipDistance,
	bLimitMax := bHardLimitMaxExceeded
			       OR bSoftLimitMaxExceeded,
	bLimitMin := bHardLimitMinExceeded
			      OR bSoftLimitMinExceeded,
	bPlusRelease := bPlusRelease,
	bMinusRelease := bMinusRelease,
	lrVelocity := SEL(NOT bReferenced, lrManualVelocity, lrVelocityNoRef),
	lrAcceleration := lrAcceleration,
	lrDeceleration := lrDeceleration,
	lrJerk := lrJerk,
	tControllerOff := tControllerOff,
	bHomeCompleted := bHomeCompleted,
	Axis := Axis,
	MasterAxis := MasterAxis
);
END_ACTION

ACTION A_AxisTerminalDiag:

(*Axis terminal diagnosis *)
fbTerminalDiagnosis(
	stTerminalState := Drive.stTerminalState,
	sTerminalStatus => sTerminalStatus
);

bErrorTerminal := NOT fbTerminalDiagnosis.bTerminalOK;
END_ACTION

END_FUNCTION_BLOCK

// ---- POUs/Tc2 Objects/Automation/Axis/Beckhoff/FB_AxisMcBeckhoffStoeberSCI6.TcPOU
FUNCTION_BLOCK FB_AxisMcBeckhoffStoeberSCI6
(*

The function block used to control axis welding.

Constructor: 		Patryk Panylo
Company:		E. Riexinger GmbH
Date:			28.04.2015
Version:			1.00

Date:			Revision:		Who:				Comment
dd.mm.yyyy		x.xx			Initials			comment

*)
VAR_INPUT
	(* Input variables / Eingang Variablen *)
	bEnable						:BOOL;						(* Axis present *)
	etMachineMode				:ET_MachineMode;			(* Machine mode *)
	etMachineState				:ET_MachineState;			(* Machine state *)
	bNoEStop					:BOOL;						(* No ermergency Stop / Keine Notaus *)
	bPowerSupplyOn				:BOOL;						(* Power supply on / Leitung eingeschaltet *)
	bLightCurtainOK				:BOOL;						(* Light curtain ok / Freigabe Lichtschranke i.o *)
	bMachineStandstill			:BOOL;						(* Machine standstill *)
	bCtrlInterrupt					:BOOL;						(* Control interrupt *)
	bMoveRelease				:BOOL;						(* Move release *)
	lrSoftLimitMax					:LREAL; 						(* Position limit switch maximum *)
	lrSoftLimitMin					:LREAL; 						(* Position limit switch minimum *)
	bTipPlus						:BOOL;						(* Manual tip in plus direction *)
	bTipMinus					:BOOL;						(* Manual tip in minus direction *)
	lrTipDistance					:LREAL;						(* Relative distance for movements *)
	bPlusRelease				:BOOL;						(* Plus move release *)
	bMinusRelease				:BOOL;						(* Minus move release *)
	bExeSetPos					:BOOL;						(* Execute set position *)
	bExeHome					:BOOL;						(* Execute home *)
	etHomingMode 				:MC_HomingMode;			(* HomingMode determines in which way the calibration is carried out. *)
	bExeMoveAbs				:BOOL;						(* Execute move absolut *)
	bExeMoveRel				:BOOL;						(* Execute move relative *)
	bExeMoveAdd				:BOOL;						(* Execute move additive *)
	bExeMoveSuper				:BOOL;						(* Execute move superimposed *)
	bExeMoveVelo				:BOOL;						(* Execute move velo *)
	bExeGearIn					:BOOL;						(* Execute gear in *)
	bExeGearOut					:BOOL;						(* Execute gear out *)
	bExeStop					:BOOL;						(* Execute move stop *)
	bExeReset					:BOOL;						(* Execute auto reset *)
	bExtOverrideEn				:BOOL;						(* External override enable *)
	lrExtOverride					:LREAL;						(* External override *)
	lrTargetPosition				:LREAL;						(* Absolute target position *)
	lrManualVelocity				:LREAL;						(* Value of velocity in manual motion [mm/s] *)
	lrVelocityNoRef				:LREAL;						(* Velocity if has no reference [mm/s] *)
	bVelocityLimitEn				:BOOL;						(* Enable velocity limit *)
	lrAutoVelocity					:LREAL;						(* Value of velocity in auto motion [mm/s] *)
	lrVelocityMin					:LREAL;						(* Velocity minimum [%] *)
	lrVelocityMax					:LREAL;						(* Velocity maximum [%] *)
	lrAcceleration					:LREAL;						(* Value of the acceleration (always positive). If >= 0 else from SM *)
	lrDeceleration				:LREAL;						(* Value of deceleration (always positive). If >= 0 else from SM *)
	lrJerk						:LREAL;						(* Value of jerk (always positive). If >= 0 else from SM *)
	bEngineTorqueLimitEn			:BOOL;						(* Enable engine torque limit *)
	lrEngineTorque				:LREAL;						(* Engine torque [%] *)
	bWithAbsoluteEncoder			:BOOL; 						(* Encoder is an absolute one / Absolutwertgeber *)
	bPosLagMonitoringEn			:BOOL;						(* Enable position lag monitoring *)
	lrOriginShiftPos				:LREAL;						(* Origin shift position *)
	dnRatioNumerator				:DINT;						(* Gear ratio numerator. Alternatively, the gear ratio can be specified in the numerator as a floating comma value, if the denominator is 1. *)
	udnRatioDenominator			:UDINT;						(* Gear ratio denominator *)
	bVeloForceCtrlEn				:BOOL;						(* Enable velocity  force controller *)
	lrVeloForceCtrlKp				:LREAL;						(* Velocity - force controller proportional band Kp *)
	lrVeloForceCtrlTi				:LREAL;						(* Velocity - force controller integral Ti *)
	lrVeloForceCtrlMin				:LREAL;						(* Velocity - force controller minimum  *)
	lrVeloForceCtrlMax			:LREAL;						(* Velocity - force controller maxmimum  *)
	lrTargetForce					:LREAL;						(* Absolute target force [N] *)
	lrForceCurrent				:LREAL;						(* Current force [mA] *)
	rForceOffset					:REAL;						(* Force offset [N] *)
	lrForceMinmA					:LREAL;						(* Force min [mA] 16#0000 = 4 [mA] *)
	lrForceMaxmA 				:LREAL;						(* Force max [mA] 16#7FFF = 20 [mA] *)
	lrForceMinN					:LREAL;						(* Force min [N] *)
	lrForceMaxN					:LREAL;						(* Force max [N] *)
	lrOverride					:LREAL;						(* Override *)
	lrActTemp					:LREAL;						(* Current temperatur *)
	lrTempLimitMax				:LREAL;						(* Temperatur limit maximum*)
	lrTempLimitMin				:LREAL;						(* Temperatur limit minimum*)
	bCoolingActive				:BOOL;						(* Cooling on *)
	snModesOfOperation			:SINT;						(* Modes of drive operation *)
	bConfirmAlarm				:BOOL;						(* Confirm alarm *)
	bOccupied					:BOOL;						(* Axis occupied *)
	tControllerOff					:TIME := t#60s;				(* Time to switch controller off *)
	tAdsTimeOut 					:TIME := t#2s;					(* Timout for ads commands *)
END_VAR
VAR_OUTPUT
	(* Output variables / Ausgang Variablen *)
	bCtrlEnabled					:BOOL;						(* Controller enabled *)
	bNotMoving					:BOOL;						(* Axis not moving *)
	bReferenced					:BOOL;						(* Axis referenced *)
	bCoupled					:BOOL;						(* Axis coupled *)
	lrActPosition					:LREAL;						(* Actual position [mm] *)
	lrActAbsPosition				:LREAL;						(* Actual absolut position [mm] *)
	lrActVelocity					:LREAL;						(* Actual velocity [mm/s] *)
	lrActForce					:LREAL;						(* Actual force [N] *)
	lrVeloMax					:LREAL;						(* Velocity limit maximum *)
	lrAccMax						:LREAL;						(* Acceleration limit maximum *)
	lrDecMax					:LREAL;						(* Deceleration limit maximum *)
	lrJerkMax					:LREAL;						(* Jerk limit maximum *)
	bHardLimitMaxExceeded		:BOOL;						(* Position limit switch maximum is exceeded *)
	bHardLimitMinExceeded		:BOOL;						(* Position limit switch minimum is exceeded *)
	bSoftLimitMaxExceeded		:BOOL;						(* Position limit switch maximum is exceeded *)
	bSoftLimitMinExceeded		:BOOL;						(* Position limit switch minimum is exceeded *)
	bCoolingOn					:BOOL;						(* Cooling *)
	bErrorTerminal				:BOOL;						(* Error Axis terminal *)
	bErrorCtrlEnabled				:BOOL;						(* Error Axis controller enabled *)
END_VAR
VAR_IN_OUT
	(* Input Output variables / Ausgang Variablen *)
	bHomeCompleted				:BOOL;						(* Home completed *)
	Drive						:ST_STOEBERSI6SC6CIA402_REF; (* The ST_STOEBERSI6SC6CIA402_REF data type  is an interface between the PLC and the DRIVE and contains axis information *)
	Axis							:AXIS_REF;					(* The AXIS_REF data type  is an interface between the PLC and the NC and contains axis information *)
	MasterAxis					:AXIS_REF;					(* The AXIS_REF data type  is an interface between the PLC and the NC and contains axis information *)
END_VAR
VAR
	(* Enummerations *)

	(* Variables *)
	sAdsAddr					:STRING(23);					(* AmsNetId of the EtherCAT master device.*)
	unSlaveAddr					:UINT;						(* Address of the slave device.*)

	nTorqueLimitMax				:INT := 100;					(* The torque limit (absolute value). Value range in %: -200 ... 200 ... 200 *)

	lrVeloLimitMax				:LREAL;
	lrVeloLimitMin					:LREAL;

	sTerminalStatus				:STRING;
	(* References *)

	(* Interfaces *)

	(* Instances *)
	fbTerminalDiagnosis			:FB_TerminalDiagnosis;
	rtMachineStandstill			:R_TRIG;
	tonAxisEnabled				:TON;

	fbController					:FB_AxisController;
	fbMoveManual				:FB_AxisMoveManual;
	fbMoveAuto					:FB_AxisMoveAuto;
	fbForce						:FB_ScalingOffset;
	fbForceCtrl					:FB_ForceController;
	fbCoolingOff					:FB_SignalHandlingDelay;
END_VAR


IF NOT bEnable								(* Signal FB enable *)
THEN

	RETURN;
END_IF

A_AxisLink();
A_AxisGetStatus();
A_AxisController();
A_AxisForceCtrl();
A_AxisMoveManual();
A_AxisMoveAuto();
A_AxisCooling();
A_AxisTerminalDiag();
A_AxisAlarm();

ACTION A_AxisAlarm:

(* Axis errors *)
tonAxisEnabled(
	IN := fbController.bEnable
		AND fbController.bRegulatorOn
		AND NOT fbController.bStatusDelay,
	PT := fbController.tStatusDelay + t#2s
);

bErrorCtrlEnabled := tonAxisEnabled.Q;
END_ACTION

ACTION A_AxisController:

(* Axis controller *)
fbController(
    	bEnable := TRUE,
	etMachineMode := etMachineMode,
	etMachineState := etMachineState,
	bRegulatorOn := bNoEStop
				      AND bPowerSupplyOn
				      AND bLightCurtainOK
				      AND SEL(bNotMoving, NOT bCtrlInterrupt, TRUE)
				      AND NOT fbMoveManual.bControllerOff
				      AND NOT fbMoveAuto.bControllerOff ,
	bReset := bConfirmAlarm,
	bTerminalOK := fbTerminalDiagnosis.bTerminalOK,
	bExeReset := bExeReset,
	bExeSetPos := bExeSetPos,
	lrSetPosition := lrTargetPosition,
	bExeGearIn := bExeGearIn,
	bExeGearOut := bExeGearOut,
	dnRatioNumerator := dnRatioNumerator,
	udnRatioDenominator := udnRatioDenominator,
	lrOverride := SEL(bExtOverrideEn,
					SEL(
						bVeloForceCtrlEn,
						lrOverride,
						fbForceCtrl.lrCVVelo),
					lrOverride*lrExtOverride/100.0),
	bWithAbsoluteEncoder := bWithAbsoluteEncoder,
	bPosLagMonitoringEn := bPosLagMonitoringEn,
	lrPositionBias := lrOriginShiftPos,
	lrSoftLimitMax := lrSoftLimitMax,
	lrSoftLimitMin := lrSoftLimitMin,
	lrAcceleration := lrAcceleration,
	lrDeceleration := lrDeceleration,
	lrJerk := lrJerk,
	Axis := Axis,
	MasterAxis := MasterAxis,
	bStatusDelay => bCtrlEnabled,
	lrActPos => lrActPosition,
	lrActAbsPos => lrActAbsPosition,
	lrActVelo => lrActVelocity,
	bNotMoving => bNotMoving,
	bReferenced => bReferenced,
	bCoupled => bCoupled,
	lrVeloLimitMax => lrVeloMax,
	lrAccLimitMax => lrAccMax,
	lrDecLimitMax => lrDecMax,
	lrJerkLimitMax => lrJerkMax,
	bHardLimitMaxExceeded => bHardLimitMaxExceeded,
	bHardLimitMinExceeded => bHardLimitMinExceeded,
	bSoftLimitMaxExceeded => bSoftLimitMaxExceeded,
	bSoftLimitMinExceeded => bSoftLimitMinExceeded
);
END_ACTION

ACTION A_AxisCooling:

(* Cooling control *)
fbCoolingOff(
	bEnable := TRUE,
	bIn := NOT bCoolingActive
		  AND lrActTemp < lrTempLimitMin
		  AND bCoolingOn,
	tDelay := t#30s
);

IF bCoolingActive
     OR lrActTemp > lrTempLimitMax
THEN
	bCoolingOn := TRUE;

ELSIF fbCoolingOff.bOut
THEN
	bCoolingOn := FALSE;
END_IF
END_ACTION

ACTION A_AxisForceCtrl:

fbForce(
	bEnable := TRUE,
	lrInput := lrForceCurrent,
	lrXLowLimit := lrForceMinmA, (* 16#0000 = 4 [mA] *)
	lrXUpperLimit := lrForceMaxmA, (* 16#7FFF = 20 [mA] *)
	lrYLowLimit := lrForceMinN,  (*[N]*)
	lrYUpperLimit := lrForceMaxN,  (*[N]*)
	usiPrecision := 2,
	lrOffset := rForceOffset,
	lrOutputPV => lrActForce
);

fbForceCtrl(
	bEnable := bNoEStop
			    AND bPowerSupplyOn
			    AND bLightCurtainOK
			    AND bCtrlEnabled,
	bControllerOn := bVeloForceCtrlEn,
	lrVeloKp := lrVeloForceCtrlKp,
	lrVeloTi := lrVeloForceCtrlTi,
	lrPVForce := lrActForce, (* [N] *)
	lrSPForce := lrTargetForce, (* [N] *)
	lrMaxForce := lrForceMaxN, (* [N] *)
	lrVeloMax := lrVeloForceCtrlMax,
	lrVeloMin := lrVeloForceCtrlMin,
	lrTaskCycle := lrgActCycleTime
);
END_ACTION

ACTION A_AxisGetStatus:

(* Get axis status *)
Axis.ReadStatus();
END_ACTION

ACTION A_AxisLink:

(* Get terminal status *)
sAdsAddr:= F_CreateAmsNetId(Drive.stTerminalState.stAdsAddr.netId);
unSlaveAddr:= Drive.stTerminalState.stAdsAddr.port;

(* Set drive parameter *)
Drive.stPlcToStoeber.snA541ModesOfOperation := snModesOfOperation;

(*Drive.PlcToStoeber.nA558TargetTorque := SEL(bEngineTorqueLimitEn,
				    nTorqueLimitMax,
				    LREAL_TO_INT(lrEngineTorque / 1.0))*)
END_ACTION

ACTION A_AxisMoveAuto:

(* Move axis auto *)
rtMachineStandstill(CLK := bMachineStandstill );

lrVeloLimitMin := SEL(bVelocityLimitEn, -1 * lrVeloMax, lrVelocityMin);
lrVeloLimitMax := SEL(bVelocityLimitEn, lrVeloMax, lrVelocityMax);

fbMoveAuto(
	bEnable := bNoEStop
               		    AND bPowerSupplyOn
               		    AND bLightCurtainOK,
	bOccupied := bOccupied,
	bCtrlEnabled := bCtrlEnabled
				      AND bMoveRelease,
	etMachineMode := etMachineMode,
	etMachineState := etMachineState,
	bReset := bConfirmAlarm,
	bExeHome := bExeHome,
	bExeMoveAbs := bExeMoveAbs,
	bExeMoveRel := bExeMoveRel,
	bExeMoveAdd := bExeMoveAdd,
	bExeMoveSuper := bExeMoveSuper,
	bExeMoveVelo := bExeMoveVelo,
	bExeStop := bExeStop
			      OR rtMachineStandstill.Q,
	etHomingMode := etHomingMode,
	lrPosition := lrTargetPosition,
	lrVelocity := LIMIT(lrVeloLimitMin, lrAutoVelocity, lrVeloLimitMax),
	lrAcceleration := lrAcceleration,
	lrDeceleration := lrDeceleration,
	lrJerk := lrJerk,
	lrOriginShiftPos := lrOriginShiftPos,
	bSignalReference := Drive.stStoeberToPlc.dwA636DigitalInputs.2,
	tControllerOff := tControllerOff,
	bHomeCompleted := bHomeCompleted,
	Axis := Axis,
	MasterAxis := MasterAxis
 );
END_ACTION

ACTION A_AxisMoveManual:

(* Move axis manual *)
fbMoveManual(
	bEnable := bNoEStop
               		    AND bPowerSupplyOn
               		    AND bLightCurtainOK,
	bOccupied := bOccupied,
	bCtrlEnabled := bCtrlEnabled
				      AND bMoveRelease,
	etMachineMode := etMachineMode,
	etMachineState := etMachineState,
	bReset := bConfirmAlarm,
	bMovePlus := bTipPlus,
	bMoveMinus := bTipMinus,
	lrTipDistance := lrTipDistance,
	bLimitMax := bHardLimitMaxExceeded
			       OR bSoftLimitMaxExceeded,
	bLimitMin := bHardLimitMinExceeded
			      OR bSoftLimitMinExceeded,
	bPlusRelease := bPlusRelease,
	bMinusRelease := bMinusRelease,
	lrVelocity := SEL(NOT bReferenced, lrManualVelocity, lrVelocityNoRef),
	lrAcceleration := lrAcceleration,
	lrDeceleration := lrDeceleration,
	lrJerk := lrJerk,
	tControllerOff := tControllerOff,
	bHomeCompleted := bHomeCompleted,
	Axis := Axis,
	MasterAxis := MasterAxis
);
END_ACTION

ACTION A_AxisTerminalDiag:

(*Axis terminal diagnosis *)
fbTerminalDiagnosis(
	stTerminalState := Drive.stTerminalState,
	sTerminalStatus => sTerminalStatus
);

bErrorTerminal := NOT fbTerminalDiagnosis.bTerminalOK;
END_ACTION

END_FUNCTION_BLOCK

// ---- POUs/Tc2 Objects/Automation/Axis/Beckhoff/FB_BECKHOFFDRIVE_REF.TcPOU
FUNCTION_BLOCK FB_BECKHOFFDRIVE_REF
VAR_INPUT
	stTerminalState			AT %I*:ST_TerminalState;
	stBECKHOFFToPlc		AT %I*:ST_BECKHOFFDRIVETOPLC;
	stPlcToBECKHOFF		AT %Q*:ST_PLCTOBECKHOFFDRIVE;
END_VAR
VAR_OUTPUT

END_VAR
VAR_IN_OUT

END_VAR
VAR

END_VAR

;

END_FUNCTION_BLOCK

// ---- POUs/Tc2 Objects/Automation/Axis/F_ChkAllAxisCoupled.TcPOU
FUNCTION F_ChkAllAxisCoupled : BOOL
(*

The function used to detect if all axis are coupled.

Constructor: 		Patryk Panylo
Company:		E. Riexinger GmbH
Date:			23.04.2015
Version:			1.00

Date:			Revision:		Who:				Comment
dd.mm.yyyy		x.xx			Initials			comment

*)
VAR_INPUT
	(* Input variables / Eingang Variablen *)
	bEnable						:BOOL;					(* Signal FB enable *)
	bAxis1Coupled				:BOOL;					(* Axis coupled *)
	bAxis2Coupled				:BOOL;					(* Axis coupled *)
	bAxis3Coupled				:BOOL;					(* Axis coupled *)
	bAxis4Coupled				:BOOL;					(* Axis coupled *)
	bAxis5Coupled				:BOOL;					(* Axis coupled *)
	bAxis6Coupled				:BOOL;					(* Axis coupled *)
	bAxis7Coupled				:BOOL;					(* Axis coupled *)
	bAxis8Coupled				:BOOL;					(* Axis coupled *)
	bAxis9Coupled				:BOOL;					(* Axis coupled *)
	bAxis10Coupled				:BOOL;					(* Axis coupled *)
END_VAR
VAR
	(* Enummerations *)

	(* Variables *)

	(* References *)

	(* Interfaces *)

	(* Instances *)

END_VAR


IF NOT bEnable							(* Signal FB enable *)
THEN
	F_ChkAllAxisCoupled := FALSE;

	RETURN;
END_IF

F_ChkAllAxisCoupled := bAxis1Coupled
					   AND bAxis2Coupled
					   AND bAxis3Coupled
					   AND bAxis4Coupled
					   AND bAxis5Coupled
					   AND bAxis6Coupled
					   AND bAxis7Coupled
					   AND bAxis8Coupled
					   AND bAxis9Coupled
					   AND bAxis10Coupled;

END_FUNCTION

// ---- POUs/Tc2 Objects/Automation/Axis/F_ChkAllAxisFieldbusOK.TcPOU
FUNCTION F_ChkAllAxisFieldbusOK : BOOL
(*

The function used to detect if all axis fieldbus ok.

Constructor: 		Patryk Panylo
Company:		E. Riexinger GmbH
Date:			23.04.2015
Version:			1.00

Date:			Revision:		Who:				Comment
dd.mm.yyyy		x.xx			Initials			comment

*)
VAR_INPUT
	(* Input variables / Eingang Variablen *)
	bEnable						:BOOL;						(* Signal FB enable *)
	bFieldbusOKAxis1				:BOOL;						(* Controller enabled *)
	bFieldbusOKAxis2				:BOOL;						(* Controller enabled *)
	bFieldbusOKAxis3				:BOOL;						(* Controller enabled *)
	bFieldbusOKAxis4				:BOOL;						(* Controller enabled *)
	bFieldbusOKAxis5				:BOOL;						(* Controller enabled *)
	bFieldbusOKAxis6				:BOOL;						(* Controller enabled *)
	bFieldbusOKAxis7				:BOOL;						(* Controller enabled *)
	bFieldbusOKAxis8				:BOOL;						(* Controller enabled *)
	bFieldbusOKAxis9				:BOOL;						(* Controller enabled *)
	bFieldbusOKAxis10			:BOOL;						(* Controller enabled *)
END_VAR
VAR
	(* Enummerations *)

	(* Variables *)

	(* References *)

	(* Interfaces *)

	(* Instances *)

END_VAR


IF NOT bEnable							(* Signal FB enable *)
THEN
	F_ChkAllAxisFieldbusOK := bEnable;

	RETURN;
END_IF

F_ChkAllAxisFieldbusOK := bFieldbusOKAxis1
					  AND bFieldbusOKAxis2
					  AND bFieldbusOKAxis3
					  AND bFieldbusOKAxis4
					  AND bFieldbusOKAxis5
					  AND bFieldbusOKAxis6
					  AND bFieldbusOKAxis7
					  AND bFieldbusOKAxis8
					  AND bFieldbusOKAxis9
					  AND bFieldbusOKAxis10;

END_FUNCTION

// ---- POUs/Tc2 Objects/Automation/Axis/F_ChkAllAxisInSamePos.TcPOU
FUNCTION F_ChkAllAxisInSamePos : BOOL
(*

The function used to detect if all axis have the same position.

Constructor: 		Patryk Panylo
Company:		E. Riexinger GmbH
Date:			09.07.2016
Version:			1.00

Date:			Revision:		Who:				Comment
dd.mm.yyyy		x.xx			Initials			comment

*)
VAR_INPUT
	(* Input variables / Eingang Variablen *)
	bEnable						:BOOL;					(* Signal FB enable *)
	lrAxis1Pos					:LREAL;					(* Axis position [mm] *)
	lrAxis2Pos					:LREAL;					(* Axis position [mm] *)
	lrAxis3Pos					:LREAL;					(* Axis position [mm] *)
	lrAxis4Pos					:LREAL;					(* Axis position [mm] *)
	lrAxis5Pos					:LREAL;					(* Axis position [mm] *)
	lrAxis6Pos					:LREAL;					(* Axis position [mm] *)
	lrAxis7Pos					:LREAL;					(* Axis position [mm] *)
	lrAxis8Pos					:LREAL;					(* Axis position [mm] *)
	lrAxis9Pos					:LREAL;					(* Axis position [mm] *)
	lrAxis10Pos					:LREAL;					(* Axis position [mm] *)
	lrTolerance					:LREAL := 2;					(* Tolerance [mm] *)
END_VAR
VAR
	(* Enummerations *)

	(* Variables *)
	nIdx1						:INT;
	nIdx2						:INT;
	arlrAxisPos					:ARRAY[1..10] OF LREAL;

	(* References *)

	(* Interfaces *)

	(* Instances *)

END_VAR


IF NOT bEnable							(* Signal FB enable *)
THEN
	F_ChkAllAxisInSamePos := TRUE;

	RETURN;
END_IF

arlrAxisPos[1] := lrAxis1Pos;
arlrAxisPos[2] := lrAxis2Pos;
arlrAxisPos[3] := lrAxis3Pos;
arlrAxisPos[4] := lrAxis4Pos;
arlrAxisPos[5] := lrAxis5Pos;
arlrAxisPos[6] := lrAxis6Pos;
arlrAxisPos[7] := lrAxis7Pos;
arlrAxisPos[8] := lrAxis8Pos;
arlrAxisPos[9] := lrAxis9Pos;
arlrAxisPos[10] := lrAxis10Pos;

F_ChkAllAxisInSamePos := TRUE;

FOR nIdx1 := 1 TO 10 DO
	FOR nIdx2 := 1 TO 10 DO
		IF ABS(arlrAxisPos[nIdx1] - arlrAxisPos[nIdx2]) > lrTolerance
		THEN
			F_ChkAllAxisInSamePos := FALSE;
			EXIT;
		END_IF
	END_FOR
END_FOR;

END_FUNCTION

// ---- POUs/Tc2 Objects/Automation/Axis/OnOff/FB_OnOff_AxisController.TcPOU
FUNCTION_BLOCK FB_OnOff_AxisController
(*

The function block used to control axis.

Constructor: 		Patryk Panylo
Company:		E. Riexinger GmbH
Date:			22.09.2015
Version:			1.00

Date:			Revision:		Who:				Comment
dd.mm.yyyy		x.xx			Initials			comment

*)
VAR_INPUT
	(* Input variables / Eingang Variablen *)
	bEnable						:BOOL;						(* Signal FB enable *)
	sAmsNetId					:STRING;					(* Ams Net Id *)
	etMachineMode				:ET_MachineMode;			(* Machine mode *)
	etMachineState				:ET_MachineState;			(* Machine state *)
	bRegulatorOn				:BOOL;						(* Enable the power stage *)
	bReset						:BOOL;						(* Signal reset *)
	bExeReset					:BOOL;						(* Execute auto reset *)
	dwRawMotorEncoder			:DWORD;					(* The raw value of the motor encoder *)
	bHWSignalLimitMax			:BOOL;						(* Signal position limit switch maximum *)
	bHWSignalLimitMin			:BOOL;						(* Signal position limit switch minimum *)
	lrSoftLimitMax					:LREAL; 						(* Position limit switch maximum *)
	lrSoftLimitMin					:LREAL; 						(* Position limit switch minimum *)
	tTimeOut 					:TIME := t#2s;					(* Timout for ads commands *)
	stEncoderConfig				:ST_EncoderConfig;			(* Encoder configuration *)
	pAxis						:POINTER TO ST_AXIS_REF_V2;				(* The AXIS_REF data type  is an interface between the PLC and the NC and contains axis information *)
END_VAR
VAR_OUTPUT
	(* Output variables / Ausgang Variablen *)
	bStatus						:BOOL;						(* Feedback *)
	bStatusDelay					:BOOL;						(* Feedback delay *)
	bError						:BOOL;						(* Controller error *)
	udnErrorNo					:UDINT;						(* Error number *)
	lrActPos						:LREAL;						(* Actual position *)
	lrActVelo						:LREAL;						(* Actual velocity *)
	bNotMoving					:BOOL;						(* Status of moving *)
	bHardLimitMaxExceeded		:BOOL;						(* Position limit switch maximum is exceeded *)
	bHardLimitMinExceeded		:BOOL;						(* Position limit switch minimum is exceeded *)
	bSoftLimitMaxExceeded		:BOOL;						(* Position limit switch maximum is exceeded *)
	bSoftLimitMinExceeded		:BOOL;						(* Position limit switch minimum is exceeded *)
END_VAR
VAR_IN_OUT

END_VAR
VAR
	(* Enummerations *)

	(* Variables *)
	tStatusDelay					:TIME := t#1s;					(* Status delay time *)
	tRegulatorOffDelay			:TIME := t#50ms;				(* Regulator off delay time *)

	bFirstTime					:BOOL;

	(* References *)

	(* Interfaces *)

	(* Instances *)
	fbPower						:FB_OnOff_Power;				(* The function block is used to enable for an axis *)
	tonStatusDelay				:TON;						(* Delay controller enabled status *)
	fbReset						:FB_OnOff_Reset;				(* An axis reset is carried out with the function block *)
	fbPositionEncoder				:FB_PositionEncoder;
END_VAR


IF NOT bEnable							(* Signal FB enable *)
THEN
	bStatus := FALSE;						(* Feedback *)
	bStatusDelay := FALSE;				(* Feedback *)
	bError := FALSE;						(* Controller error *)
	udnErrorNo := 0;						(* Error number *)

	bFirstTime := FALSE;
	RETURN;
END_IF

IF NOT bFirstTime
THEN

	bFirstTime := TRUE;
END_IF;

A_MCPower();
A_MCReset();
A_PositionDynamics();
A_GetLimits();
A_SetLimits();
A_Error();

(* Actual position *)
lrActPos := pAxis^.stPosition.lrActPos;
lrActPos := F_LRealRound(lrReal := lrActPos, usiPrecision := 2);

(* Actual velocity *)
lrActVelo := pAxis^.stDynamics.lrActVelo;
lrActVelo := F_LRealRound(lrReal := lrActVelo, usiPrecision := 2);

(* Current engine torque *)
(*nActEngineTorque := Axis.stNcToPlc.nActEngineTorque;*)

(* Status not moving *)
bNotMoving := NOT pAxis^.stAxisStates.bOperational                          		(* Control enabled *)
			  OR pAxis^.stAxisStates.bNotMoving;					(* Axis standstill *)

ACTION A_Error:

bError := fbReset.bError
	         OR fbPower.bError;
END_ACTION

ACTION A_GetLimits:

(* Status hardware limit switch *)
bHardLimitMaxExceeded := pAxis^.stLimitSwitches.bHWLimitMax;						(* Position limit switch maximum is exceeded *)
bHardLimitMinExceeded := pAxis^.stLimitSwitches.bHWLimitMin;						(* Position limit switch minimum is exceeded *)

(* Status software limit switch *)
bSoftLimitMaxExceeded := lrActPos >= lrSoftLimitMax;			(* Position limit switch maximum is exceeded *)
bSoftLimitMinExceeded := lrActPos <= lrSoftLimitMin;			(* Position limit switch minimum is exceeded *)


pAxis^.stLimitSwitches.lrSWPosLimitMax := lrSoftLimitMax;
pAxis^.stLimitSwitches.lrSWPosLimitMin := lrSoftLimitMin;
pAxis^.stLimitSwitches.bSWLimitMaxActive := bSoftLimitMaxExceeded;
pAxis^.stLimitSwitches.bSWLimitMinActive := bSoftLimitMinExceeded;
END_ACTION

ACTION A_MCPower:

fbPower(
	bEnable := TRUE,
	bRegulatorOn := bRegulatorOn,
	bEnablePositive := bHWSignalLimitMax,                         			(* HW limit switch maximum *)
	bEnableNegative := bHWSignalLimitMin,                         			(* HW Limit switch minimum *)
	pAxis := pAxis,
	bStatus => bStatus
);

tonStatusDelay(
	IN := fbPower.bStatus,
	PT := SEL(etMachineMode = ET_MachineMode_eManual, tStatusDelay, t#0ms),
	Q => bStatusDelay
);
END_ACTION

ACTION A_MCReset:

fbReset(
	bExecute := bReset
	            	     XOR bExeReset,
	pAxis := pAxis
);
END_ACTION

ACTION A_PositionDynamics:

(* Position encoding *)
fbPositionEncoder(
	bEnable := TRUE,
	dwEncCurrentValue := dwRawMotorEncoder,
	stEncCfg := stEncoderConfig,
	pAxis := pAxis
);
END_ACTION

ACTION A_SetLimits:

;
END_ACTION

END_FUNCTION_BLOCK

// ---- POUs/Tc2 Objects/Automation/Axis/OnOff/FB_OnOff_AxisMoveAuto.TcPOU
FUNCTION_BLOCK FB_OnOff_AxisMoveAuto
(*

The function block used to auto control of axis.

Constructor: 		Patryk Panylo
Company:		E. Riexinger GmbH
Date:			22.09.2015
Version:			1.00

Date:			Revision:		Who:				Comment
dd.mm.yyyy		x.xx			Initials			comment

*)
VAR_INPUT
	(* Input variables / Eingang Variablen *)
	bEnable						:BOOL;						(* Signal FB enable *)
	etMachineMode				:ET_MachineMode;			(* Machine mode *)
	etMachineState				:ET_MachineState;			(* Machine state *)
	bCtrlEnabled					:BOOL;						(* Controller enabled *)
	bReset						:BOOL;						(* Reset *)
	bExeMoveAbs				:BOOL;						(* Execute move absolut *)
	bSuperImposedOn			:BOOL;						(* Switch SuperImposed on / off *)
	bExeMoveVelo				:BOOL;						(* Execute move velo *)
	bExeStop					:BOOL;						(* Execute stop *)
	lrPosition						:LREAL;						(* Target position *)
	lrVelocity						:LREAL;						(* Target velocity *)
	tControllerOff					:TIME := t#60s;				(* Time to switch controller off *)
	stControllerConfig				:ST_VeloControllerConfig;				(* Controller configuration *)
	pAxis						:POINTER TO ST_AXIS_REF_V2;				(* The AXIS_REF data type  is an interface between the PLC and the NC and contains axis information *)
END_VAR
VAR_OUTPUT
	(* Output variables / Ausgang Variablen *)
	bInPosition					:BOOL;						(* Target position is reached *)
	bInVelocity					:BOOL;						(* Target velocity is reached *)
	bStopped					:BOOL;						(* Target stopped *)
	bControllerOff					:BOOL;						(* Switch controller off *)
	bMoveToPlus				:BOOL;						(* Move to plus *)
	bMoveToMinus				:BOOL;						(* Move to minus *)
	bError						:BOOL;						(* Program error *)
	udnErrorNo					:UDINT;						(* Error number *)
END_VAR
VAR_IN_OUT
	bHomeCompleted				:BOOL;						(* Home completed *)
END_VAR
VAR
	(* Enummerations *)

	(* Variables *)

	bFirstTime					:BOOL;

	(* References *)

	(* Interfaces *)

	(* Instances *)
	fbMoveAbs					:FB_OnOff_MoveAbsolut;
	fbMoveVelo					:FB_OnOff_MoveVelocity;
	fbStop						:FB_OnOff_Stop;
	fbPositionController			:FB_PositionController;
	fbStateIdle					:FB_SignalWatchdog;
END_VAR


IF NOT bEnable								(* Signal FB enable *)
THEN
	(* The function block MoveAbsolute starts positioning to an absolute target position and monitors the axis movement over the whole travel path.  *)
	fbMoveAbs(
		bExecute := FALSE,
		pAxis := pAxis,
		bDone => bInPosition
	);

	(* The function block MoveVelocity starts a continuous movement with specified velocity and direction.  *)
	fbMoveVelo(
		bExecute := FALSE,
		pAxis := pAxis,
		bInVelocity => bInVelocity
	 );

	(* The function block Stop stops an axis with a defined braking ramp and blocks the axis for any motion commands.  *)
	fbStop(
		bExecute := FALSE,
		pAxis := pAxis,
		bDone => bStopped
	);

	fbStateIdle(
		bEnable := FALSE,
		tWatchdog := tControllerOff
	);

	bMoveToPlus := FALSE;
	bMoveToMinus := FALSE;

	bControllerOff := FALSE;

	bFirstTime := FALSE;

	RETURN;
END_IF;

IF NOT bFirstTime
THEN

	bFirstTime := TRUE;
END_IF;

IF bReset
     AND bError
THEN
	(* The function block MoveAbsolute starts positioning to an absolute target position and monitors the axis movement over the whole travel path.  *)
	fbMoveAbs(
		bExecute := FALSE,
		pAxis := pAxis,
		bDone => bInPosition
	);

	(* The function block MoveVelocity starts a continuous movement with specified velocity and direction.  *)
	fbMoveVelo(
		bExecute := FALSE,
		pAxis := pAxis,
		bInVelocity => bInVelocity
	 );

	(* The function block Stop stops an axis with a defined braking ramp and blocks the axis for any motion commands.  *)
	fbStop(
		bExecute := FALSE,
		pAxis := pAxis,
		bDone => bStopped
	);

	bMoveToPlus := FALSE;
	bMoveToMinus := FALSE;
END_IF;

IF bCtrlEnabled
     AND (etMachineMode = ET_MachineMode_eAutomatic
		OR etMachineMode = ET_MachineMode_eStepping
		OR etMachineMode = ET_MachineMode_eHome)
    AND etMachineState <> ET_MachineState_eIdle
    AND etMachineState <> ET_MachineState_eUndefined
THEN
	(* The function block MoveAbsolute starts positioning to an absolute target position and monitors the axis movement over the whole travel path.  *)
	fbMoveAbs(
		bExecute := bExeMoveAbs,
		lrPosition := lrPosition,
		bSuperImposed := bSuperImposedOn,
		pAxis := pAxis,
		bDone => bInPosition
	);

	(* The function block MoveVelocity starts a continuous movement with specified velocity and direction.  *)
	fbMoveVelo(
		bExecute := bExeMoveVelo,
		lrVelocity	 := lrVelocity,
		pAxis := pAxis,
		bInVelocity => bInVelocity
	 );

	A_Controller();

	pAxis^.stPosition.lrSetPos := LIMIT(
		pAxis^.stLimitSwitches.lrSWPosLimitMin,
		pAxis^.stPosition.lrSetPos ,
		pAxis^.stLimitSwitches.lrSWPosLimitMax
	);

	bMoveToPlus := NOT pAxis^.stAxisCtrl.bQuickStop
				      AND (fbMoveAbs.bMoveToPlus
						OR fbMoveVelo.bMoveToPlus);

	bMoveToMinus := NOT pAxis^.stAxisCtrl.bQuickStop
				         AND (fbMoveAbs.bMoveToMinus
						   OR fbMoveVelo.bMoveToMinus);

ELSE
	(* The function block MoveAbsolute starts positioning to an absolute target position and monitors the axis movement over the whole travel path.  *)
	fbMoveAbs(
		bExecute := FALSE,
		pAxis := pAxis,
		bDone => bInPosition
	);

	(* The function block MoveVelocity starts a continuous movement with specified velocity and direction.  *)
	fbMoveVelo(
		bExecute := FALSE,
		pAxis := pAxis,
		bInVelocity => bInVelocity
	 );

	bMoveToPlus := FALSE;
	bMoveToMinus := FALSE;

END_IF;

fbStateIdle(
	bEnable := etMachineMode = ET_MachineMode_eAutomatic
			    OR etMachineMode = ET_MachineMode_eStepping
		  	    OR etMachineMode = ET_MachineMode_eHome,
	bIn := etMachineState <> ET_MachineState_eIdle
		  AND etMachineState <> ET_MachineState_eUndefined,
	tWatchdog := tControllerOff
);

bControllerOff := NOT fbStateIdle.bOut
			    AND (etMachineMode = ET_MachineMode_eAutomatic
				        OR etMachineMode = ET_MachineMode_eStepping
				        OR etMachineMode = ET_MachineMode_eHome);

(* The function block Stop stops an axis with a defined braking ramp and blocks the axis for any motion commands.  *)
fbStop(
	bExecute := bExeStop,
	pAxis := pAxis,
	bDone => bStopped
);

pAxis^.stAxisStates.bNotMoving := NOT bMoveToPlus
							    AND NOT bMoveToMinus;

bError :=  fbMoveAbs.bError
		OR fbMoveVelo.bError
		OR fbStop.bError;

ACTION A_Controller:

fbPositionController (
	bEnable := TRUE,
	dnSetPos := pAxis^.stPosition.dnSetPos,
	stCtrlCfg := stControllerConfig,
(*	lrPosMin := ,
	lrPosMax := ,*)
	pAxis := pAxis,
	lrVeloOut => ,
	lrProcessErr => ,
	bVeloMin => ,
	bVeloMax =>
);
END_ACTION

END_FUNCTION_BLOCK

// ---- POUs/Tc2 Objects/Automation/Axis/OnOff/FB_OnOff_AxisMoveManual.TcPOU
FUNCTION_BLOCK FB_OnOff_AxisMoveManual
(*

The function block used to manual control of axis.

Constructor: 		Patryk Panylo
Company:		E. Riexinger GmbH
Date:			22.09.2015
Version:			1.00

Date:			Revision:		Who:				Comment
dd.mm.yyyy		x.xx			Initials			comment

*)
VAR_INPUT
	(* Input variables / Eingang Variablen *)
	bEnable						:BOOL;						(* Signal FB enable *)
	etMachineMode				:ET_MachineMode;			(* Machine mode *)
	etMachineState				:ET_MachineState;			(* Machine state *)
	bNoEStop					:BOOL;						(* No ermergency Stop / Keine Notaus *)
	bPowerSupplyOn				:BOOL;						(* Power supply on / Leitung eingeschaltet *)
	bLightCurtainOK				:BOOL;						(* Light curtain ok / Freigabe Lichtschranke i.o *)
	bReset						:BOOL;						(* Reset *)
	bMovePlus					:BOOL;						(* Move in plus direction *)
	bMoveMinus					:BOOL;						(* Move in minus direction *)
	bInPlusLimit					:BOOL;						(* In plus limit *)
	bInMinusLimit					:BOOL;						(* In minus limit *)
	bPlusRelease				:BOOL;						(* Plus move release *)
	bMinusRelease				:BOOL;						(* Minus move release *)
	tTimeOut						:TIME := t#5s;					(* TimeOut *)
END_VAR
VAR_OUTPUT
	(* Output variables / Ausgang Variablen *)
	bMoving						:BOOL;						(* Axis moving *)
	bMoveToPlus				:BOOL;						(* Move to plus *)
	bMoveToMinus				:BOOL;						(* Move to minus *)
	bErrorMoveToPlus			:BOOL;						(* Error move to plus *)
	bErrorMoveToMinus			:BOOL;						(* Error move to minus *)
END_VAR
VAR_IN_OUT
	bHomeCompleted				:BOOL;						(* Home completed *)
END_VAR
VAR
	(* Enummerations *)

	(* Variables *)
	bFirstTime					:BOOL;

	(* References *)

	(* Interfaces *)

	(* Instances *)
	fbJog						:FB_Motor;					(* The function block is used to manual control an axis *)
	fbAtPlusLimit					:FB_SignalHandlingDelay;
	fbAtMinusLimit				:FB_SignalHandlingDelay;
	fbPlusRelease				:FB_SignalHandlingDelay;
	fbMinusRelease				:FB_SignalHandlingDelay;
END_VAR


IF NOT bEnable							(* Signal FB enable *)
THEN
	fbJog(
		bEnable := FALSE,
		bHandPlus := FALSE,
		bHandMinus := FALSE,
		bAutoPlus := FALSE,
		bAutoMinus := FALSE,
		bHomeCompleted := bHomeCompleted,
		bMoveToPlus => bMoveToPlus,
		bMoveToMinus => bMoveToMinus
	);

	bFirstTime := FALSE;

	RETURN;
END_IF

IF NOT bFirstTime
THEN

	bFirstTime := TRUE;
END_IF

(* Control on/off motor *)
fbAtPlusLimit(
	bEnable := TRUE,
	bIn := bInPlusLimit,
	tDelay := t#0ms
);

fbAtMinusLimit(
	bEnable := TRUE,
	bIn := bInMinusLimit,
	tDelay := t#0ms
);

fbPlusRelease(
	bEnable := TRUE,
	bIn := bPlusRelease,
	tDelay :=t#0ms
);

fbMinusRelease(
	bEnable := TRUE,
	bIn := bMinusRelease,
	tDelay := t#0ms
);

fbJog(
	bEnable := TRUE,
	bNoEmergencyStop := bNoEStop
						AND bLightCurtainOK,
	bVoltageOK := bPowerSupplyOn,
	bReset := bReset,
	bAutoHand := etMachineMode = ET_MachineMode_eHome
			         OR etMachineMode = ET_MachineMode_eStepping
			         OR etMachineMode = ET_MachineMode_eAutomatic,
	bHandPlus := bMovePlus,
	bHandMinus := bMoveMinus,
	bAtPlusLimit := fbAtPlusLimit.bOut,
	bAtMinusLimit := fbAtMinusLimit.bOut,
	bPlusRelease := fbPlusRelease.bOut,
	bMinusRelease := fbMinusRelease.bOut,
	bSyncPlus := FALSE,
	bSyncMinus := FALSE,
	bSyncOn := FALSE,
	bControlOff := FALSE,
	bMotorCtrlErrOff := FALSE,
	bErrorOff := TRUE,
	tSyncTimeOut := ,
	tConTimeOut := ,
	tCtrlTimeOut := tTimeOut,
	bHomeCompleted := bHomeCompleted,
	bMoveToPlus => bMoveToPlus,
	bMoveToMinus => bMoveToMinus
);

A_Error();

ACTION A_Error:

bErrorMoveToMinus := fbJog.bError
					AND (fbJog.udnErrorNo = 1
					     OR fbJog.udnErrorNo = 2
					     OR fbJog.udnErrorNo = 5);

bErrorMoveToPlus := fbJog.bError
					 AND (fbJog.udnErrorNo = 3
					       OR fbJog.udnErrorNo = 4
					       OR fbJog.udnErrorNo = 5);
END_ACTION

END_FUNCTION_BLOCK

// ---- POUs/Tc2 Objects/Automation/Axis/VFD/FB_VFD_AxisController.TcPOU
FUNCTION_BLOCK FB_VFD_AxisController
(*

The function block used to control drive.

Constructor: 		Patryk Panylo
Company:		E. Riexinger GmbH
Date:			14.06.2018
Version:			1.00

Date:			Revision:		Who:				Comment
dd.mm.yyyy		x.xx			Initials			comment

*)
VAR_INPUT
	(* Input variables / Eingang Variablen *)
	bEnable						:BOOL;						(* Signal FB enable *)
	etMachineMode				:ET_MachineMode;			(* Machine mode *)
	etMachineState				:ET_MachineState;			(* Machine state *)
	bRegulatorOn				:BOOL;						(* Enable the controller stage *)
	bReset						:BOOL;						(* Signal reset *)
	bExeReset					:BOOL;						(* Execute auto reset *)
	lrOverride					:LREAL;						(* Override 100% percent *)
END_VAR
VAR_OUTPUT
	(* Output variables / Ausgang Variablen *)
	bStatus						:BOOL;						(* Feedback *)
	bStatusDelay					:BOOL;						(* Feedback delay *)
	lrActVelo						:LREAL;						(* Actual velocity *)
	bNotMoving					:BOOL;						(* Status of moving *)
	bError						:BOOL;						(* Controller error *)
	bErrorInit						:BOOL;						(* Controller initialization error *)
	udnErrorNo					:UDINT;						(* Error number *)
END_VAR
VAR_IN_OUT
	Axis							:ST_VFD_AXIS_REF;			(* The AXIS_REF data type  is an interface between the PLC and the NC and contains axis information *)
END_VAR
VAR
	(* Enummerations *)

	(* Variables *)
	tStatusDelay					:TIME := t#1s;					(* Status delay time *)
	tRegulatorOffDelay			:TIME := t#50ms;				(* Regulator off delay time *)

	bFirstTime					:BOOL;

	(* References *)

	(* Interfaces *)

	(* Instances *)
	fbPower						:FB_VFD_Power;			(* The function block is used to enable for an drive *)
	tonStatusDelay				:TON;					(* Delay controller enabled status *)
	fbReset						:FB_VFD_Reset;			(* An drive reset is carried out with the function block *)

END_VAR


IF NOT bEnable							(* Signal FB enable *)
THEN
	bStatus := FALSE;						(* Feedback *)
	bStatusDelay := FALSE;				(* Feedback *)
	bError := FALSE;						(* Controller error *)
	udnErrorNo := 0;						(* Error number *)

	bNotMoving := TRUE;
	lrActVelo := 0;

	bFirstTime := FALSE;
	RETURN;
END_IF

IF NOT bFirstTime
THEN

	bFirstTime := TRUE;
END_IF;

A_Power();
A_Reset();
A_Error();

(* Status not moving *)
bNotMoving := Axis.bNotMoving;					(* Drive standstill *)

(* Actual velocity *)
lrActVelo := INT_TO_LREAL(Axis.nCurrentMotorSpeed) * (24000.0/32767.0);
lrActVelo := F_LRealRound(lrReal := lrActVelo, usiPrecision := 2);

ACTION A_Error:

bError := fbReset.bError
	         OR fbPower.bError;

bErrorInit := FALSE;
END_ACTION

ACTION A_Power:

fbPower(
	bEnable := TRUE,
	bRegulatorOn := bRegulatorOn,
	lrOverride := lrOverride,
	Axis := Axis,
	bStatus => bStatus
);

tonStatusDelay(
	IN := fbPower.bStatus,
	PT := SEL(etMachineMode = ET_MachineMode_eManual, tStatusDelay, t#0ms),
	Q => bStatusDelay
);
END_ACTION

ACTION A_Reset:

fbReset(
	bExecute := bReset
	            	     XOR bExeReset,
	Axis := Axis
);
END_ACTION

END_FUNCTION_BLOCK

// ---- POUs/Tc2 Objects/Automation/Axis/VFD/FB_VFD_AxisLink.TcPOU
FUNCTION_BLOCK FB_VFD_AxisLink
VAR_INPUT
END_VAR
VAR_OUTPUT
END_VAR
VAR_IN_OUT
	Drive						:ST_VFD_DRIVE_REF;			(* The DRIVE_REF data type  is an interface between the PLC and the DRIVE and contains axis information *)
	Axis							:ST_VFD_AXIS_REF;			(* The AXIS_REF data type  is an interface between the PLC and the NC and contains axis information *)
END_VAR
VAR

END_VAR
VAR CONSTANT
	rAxFactor		:REAL := 0.9328;
	rBFactor			:REAL := 98.0;
END_VAR


(* Set terminal parameters *)
Axis.sAdsAddr:= F_CreateAmsNetId(Drive.stTerminalState.stAdsAddr.netId);
Axis.unSlaveAddr:= Drive.stTerminalState.stAdsAddr.port;

(* Copy the actual values from the inverter to the axis reference *)
Axis.bEnabled := Drive.stVfdToPlc.bEnabled;										(* The drive is enabled. *)
Axis.bOperational := Drive.stVfdToPlc.bOperational OR Drive.stVfdToPlc.bEnabled;		(* The drive is ready for operation. *)
Axis.bError := Drive.stVfdToPlc.bBrakeError OR NOT Drive.stVfdToPlc.bEnabled;		(* The drive state is fault. *)
Axis.bNotMoving := Drive.stVfdToPlc.nCurrentMotorSpeed < 50;						(* Motor not moving *)
Axis.bMotorSpeedReached := Axis.nSetMotorSpeed > 50								(* Motor speed reached *)
						     AND (ABS(Axis.nCurrentMotorSpeed - Axis.nSetMotorSpeed) < 100);
Axis.nCurrentMotorSpeed := REAL_TO_INT((Drive.stVfdToPlc.nCurrentMotorSpeed * rAxFactor) + rBFactor);					(* Current motor speed *)

(* Copy the setpoint values from the axis reference to the inverter *)
Drive.stPlcToVfd.bEnable := Axis.bEnable;										(* Enable controller *)
Drive.stPlcToVfd.bFaultReset := Axis.bFaultReset;									(* Acknowledgment for faults of the device state machine. *)
Drive.stPlcToVfd.bForwardStop:= Axis.bForwardStop;								(* Counterclockwise rotation moving. *)
Drive.stPlcToVfd.bReverseStop:= Axis.bReverseStop;								(* Clockwise rotation moving. *)
Drive.stPlcToVfd.bJog:= Axis.bJog;												(* Jog command. *)
Drive.stPlcToVfd.bExtError:= Axis.bExtError;										(* External error signal. *)
Drive.stPlcToVfd.nSetMotorSpeed := Axis.nSetMotorSpeed * (Axis.nOverride/100) ;	(* Relative speed reference value *)
Drive.stPlcToVfd.bReserve1 := Axis.bReserve1;									(* Reserve 1. *)
Drive.stPlcToVfd.bReserve2 := Axis.bReserve2;									(* Reserve 2. *)

END_FUNCTION_BLOCK

// ---- POUs/Tc2 Objects/Automation/Axis/VFD/FB_VFD_AxisMoveAuto.TcPOU
FUNCTION_BLOCK FB_VFD_AxisMoveAuto
(*

The function block used to auto control of axis.

Constructor: 		Patryk Panylo
Company:		E. Riexinger GmbH
Date:			14.06.2018
Version:			1.00

Date:			Revision:		Who:				Comment
dd.mm.yyyy		x.xx			Initials			comment

*)
VAR_INPUT
	(* Input variables / Eingang Variablen *)
	bEnable						:BOOL;						(* Signal FB enable *)
	etMachineMode				:ET_MachineMode;			(* Machine mode *)
	etMachineState				:ET_MachineState;			(* Machine state *)
	bCtrlEnabled					:BOOL;						(* Controller enabled *)
	bReset						:BOOL;						(* Reset *)
	bExeMoveVelo				:BOOL;						(* Execute move velo *)
	bExeStop					:BOOL;						(* Execute stop *)
	lrVelocity						:LREAL;						(* Target velocity *)
	lrSpeedLimitMax				:LREAL;						(* Maximal speed *)
	tControllerOff					:TIME := t#60s;				(* Time to switch controller off *)
END_VAR
VAR_OUTPUT
	(* Output variables / Ausgang Variablen *)
	bInVelocity					:BOOL;						(* Target velocity is reached *)
	bStopped					:BOOL;						(* Target stopped *)
	bControllerOff					:BOOL;						(* Switch controller off *)
	bError						:BOOL;						(* Program error *)
	udnErrorNo					:UDINT;						(* Error number *)
END_VAR
VAR_IN_OUT
	bHomeCompleted				:BOOL;						(* Home completed *)
	Axis							:ST_VFD_AXIS_REF;			(* The AXIS_REF data type  is an interface between the PLC and the NC and contains axis information *)
END_VAR
VAR
	(* Enummerations *)

	(* Variables *)

	bFirstTime					:BOOL;

	(* References *)

	(* Interfaces *)

	(* Instances *)
	fbMoveVelo					:FB_VFD_MoveVelocity;
	fbStop						:FB_VFD_Stop;
	fbStateIdle					:FB_SignalWatchdog;
END_VAR


IF NOT bEnable								(* Signal FB enable *)
THEN
	(* The function block MoveVelocity starts a continuous movement with specified velocity and direction.  *)
	fbMoveVelo(
		bExecute := FALSE,
		Axis := Axis,
		bInVelocity => bInVelocity
	 );

	(* The function block Stop stops an axis with a defined braking ramp and blocks the axis for any motion commands.  *)
	fbStop(
		bExecute := FALSE,
		Axis := Axis,
		bDone => bStopped
	);

	fbStateIdle(
		bEnable := FALSE,
		tWatchdog := tControllerOff
	);

	bControllerOff := FALSE;

	bFirstTime := FALSE;

	RETURN;
END_IF;

IF NOT bFirstTime
THEN

	bFirstTime := TRUE;
END_IF;

IF bReset
     AND bError
THEN
	(* The function block MoveVelocity starts a continuous movement with specified velocity and direction.  *)
	fbMoveVelo(
		bExecute := FALSE,
		Axis := Axis,
		bInVelocity => bInVelocity
	 );

	(* The function block Stop stops an axis with a defined braking ramp and blocks the axis for any motion commands.  *)
	fbStop(
		bExecute := FALSE,
		Axis := Axis,
		bDone => bStopped
	);

END_IF;

IF bCtrlEnabled
     AND (etMachineMode = ET_MachineMode_eAutomatic
		OR etMachineMode = ET_MachineMode_eStepping
		OR etMachineMode = ET_MachineMode_eHome)
    AND etMachineState <> ET_MachineState_eIdle
    AND etMachineState <> ET_MachineState_eUndefined
THEN
	(* The function block MoveVelocity starts a continuous movement with specified velocity and direction.  *)
	fbMoveVelo(
		bExecute := bExeMoveVelo,
		lrVelocity	 := lrVelocity,
		lrVelocityMax := lrSpeedLimitMax,
		Axis := Axis,
		bInVelocity => bInVelocity
	 );

ELSE
	(* The function block MoveVelocity starts a continuous movement with specified velocity and direction.  *)
	fbMoveVelo(
		bExecute := FALSE,
		Axis := Axis,
		bInVelocity => bInVelocity
	 );

END_IF;

fbStateIdle(
	bEnable := etMachineMode = ET_MachineMode_eAutomatic
			    OR etMachineMode = ET_MachineMode_eStepping
		  	    OR etMachineMode = ET_MachineMode_eHome,
	bIn := etMachineState <> ET_MachineState_eIdle
		  AND etMachineState <> ET_MachineState_eUndefined,
	tWatchdog := tControllerOff
);

bControllerOff := NOT fbStateIdle.bOut
			    AND (etMachineMode = ET_MachineMode_eAutomatic
				        OR etMachineMode = ET_MachineMode_eStepping
				        OR etMachineMode = ET_MachineMode_eHome);

(* The function block Stop stops an axis with a defined braking ramp and blocks the axis for any motion commands.  *)
fbStop(
	bExecute := bExeStop,
	Axis := Axis,
	bDone => bStopped
);

A_Error();

ACTION A_Error:

bError := fbMoveVelo.bError
	        OR fbStop.bError;
END_ACTION

END_FUNCTION_BLOCK

// ---- POUs/Tc2 Objects/Automation/Extraction Fan/FB_ExtractionFan.TcPOU
FUNCTION_BLOCK FB_ExtractionFan
(*

The function block used to control extraction fan.

Constructor: 		Patryk Panylo
Company:		E. Riexinger GmbH
Date:			07.09.2018
Version:			1.00

Date:			Revision:		Who:				Comment
xx.xx.xxxx			1.01									

*)
VAR_INPUT
	(* Input variables / Eingang Variablen *)
	bEnable							:BOOL;						(* Function block enable *)
	bNoEStop						:BOOL;						(* No ermergency Stop / Keine Notaus *)
	bPowerSupplyOn					:BOOL;						(* Power supply on / Leitung eingeschaltet *)
	bLightCurtainOK					:BOOL;						(* Light curtain ok / Freigabe Lichtschranke i.o *)
	bReset							:BOOL;						(* Controller reset *)
	bAutoHand						:BOOL;						(* Auto := TRUE, Hand := FALSE *)
	bHandOn						:BOOL;						(* Heater on/off in manual mode with rising edge *)
	bAutoOn							:BOOL;						(* Heater on/off in auto mode rising edge *)
	bAutoOff							:BOOL;						(* Heater off in auto mode with rising edge *)
	bReleaseOn						:BOOL;						(* Release on *)
	bCtrlInterrupt						:BOOL;						(* Control interrupt *)
	lrSPPower						:LREAL;						(* Setpoint of power 0 - 100 % *)
	bEnAutoCtrlOff					:BOOL := FALSE;				(* Auto off enable*)
	tCtrlPowerOff						:TIME := t#90s;				(* Time to switch controller power off *)
	tCtrlPowerOn						:TIME := t#90s;				(* Time to switch controller power on *)
	lrPowerMin						:LREAL;						(* Power minimum *)
	lrPowerMax						:LREAL;						(* Power maximum *)
	lrSetTemp						:LREAL;						(* Set temperature *)
	lrActTemp						:LREAL;						(* Actual temperature *)
	lrMaxTemp						:LREAL;						(* Maximal temperature *)
	tReadyDelay						:TIME := T#5s;				(* Ready delay*)
	tTimeOut							:TIME := T#5s;				(* TimeOut *)
END_VAR
VAR_OUTPUT
	(* Output variables / Ausgang Variablen *)
	bPowerOn						:BOOL;						(* Power on *)
	unCVPower						:UINT;						(* Current value of power 0 - 10 V *)
	bReady 							:BOOL;						(* Heater ready *)
	bError							:BOOL;						(* Program error  *)
	udnErrorNo						:UDINT;						(* Error number *)
	sErrorMsg						:STRING; 					(* Error message *)
END_VAR
VAR_IN_OUT
	(* Input Output variables / Ausgang Variablen *)

END_VAR
VAR
	(* Enummerations *)

	(* Variables *)
	bReleasePowerOn				:BOOL;

	bFirstTime						:BOOL;

	(* References *)

	(* Interfaces *)

	(* Instances *)
	tonWatchDog						:TON;
	tonPowerSupplyOn				:TON;
	fbCtrlPowerOff					:FB_SignalHandlingDelay;
	fbCtrlPowerOn					:FB_SignalHandlingDelay;
	fbScalingSP						:FB_Scaling;
	fbReadyDelay					:FB_SignalHandlingDelay;

	rtHandOn						:R_TRIG;
	rtAutoOn							:R_TRIG;
	rtAutoOff							:R_TRIG;
END_VAR
VAR CONSTANT

END_VAR


IF NOT bEnable
THEN
	bPowerOn := FALSE;				(* Power on *)
 	unCVPower := 0;					(* Current value of power 0 - 100 % *)
	bReady := TRUE;				(* Heater enabled *)
	bError := FALSE;					(* Program error  *)
	udnErrorNo := 0;					(* Error number *)
	sErrorMsg := ''; 					(* Error message *)
	tonWatchDog(IN := FALSE);

	bFirstTime := FALSE;
	RETURN;
END_IF

IF NOT bFirstTime
THEN
	bReleasePowerOn := TRUE;

	bPowerOn := FALSE;				(* Powr on *)
 	unCVPower := 0;					(* Current value of power 0 - 100 % *)
	bReady := FALSE;				(* Heater enabled *)

	bFirstTime := TRUE;
END_IF

(* Controller automatic off *)
fbCtrlPowerOff(
	bEnable := TRUE,
	bIn := bEnAutoCtrlOff
		  AND bAutoHand					(* Automatic *)
		  AND bPowerOn,
	tDelay := tCtrlPowerOff
);

fbCtrlPowerOn(
	bEnable := TRUE,
	bIn := NOT bPowerOn					(* Ctrl disabled *)
		  AND NOT bReleasePowerOn,
	tDelay := tCtrlPowerOn
);

IF NOT bNoEStop
     OR NOT bPowerSupplyOn
     OR NOT bLightCurtainOK
     OR bError
     OR bCtrlInterrupt
     OR fbCtrlPowerOff.bOut
THEN
	bReleasePowerOn := FALSE;
	bPowerOn := FALSE;

ELSIF fbCtrlPowerOn.bOut
THEN
	bReleasePowerOn := TRUE;
END_IF

IF bReset
     AND bError
THEN
	udnErrorNo := 0;					(* Error number *)
	sErrorMsg := ''; 					(* Error message *)
	tonWatchDog(IN := FALSE);

END_IF

(* Check inputs  *)
rtHandOn(CLK := bHandOn);
rtAutoOn(CLK := bAutoOn AND bReleaseOn AND bReleasePowerOn);
rtAutoOff(CLK := bAutoOff);

(* Check operating mode *)
IF bAutoHand					(* Automatic *)
THEN
	IF rtAutoOff.Q
	THEN
		bPowerOn := FALSE;

	ELSIF rtAutoOn.Q
		    AND bReleasePowerOn
	THEN
		bPowerOn := TRUE;

		fbCtrlPowerOff(bEnable := FALSE);
		fbCtrlPowerOn(bEnable := FALSE);
	END_IF;

ELSE						(* Manual *)
	IF rtHandOn.Q
	THEN
		IF bPowerOn
		THEN
			bPowerOn := FALSE;

		ELSIF bReleaseOn
			   AND bReleasePowerOn
		THEN
			bPowerOn := TRUE;
		END_IF
	END_IF

END_IF;

(* Timer starts when cylinder is not  in base and work position *)
tonWatchDog(
	IN := bPowerOn
		 AND bPowerSupplyOn
		 AND NOT bReady,
	PT := SEL(bAutoHand, tTimeOut, tTimeOut + tReadyDelay)
);

(* Error if cylinder does not reach base or work position*)
IF tonWatchDog.Q
   AND NOT bError
THEN
	IF bPowerOn AND NOT bReady
	THEN
		udnErrorNo := 1; 								(* Set error number *)
		sErrorMsg := 'Not ready error';
	END_IF
END_IF

tonPowerSupplyOn(
	IN := bNoEStop
		AND NOT bPowerSupplyOn,
	PT := t#3s
);

IF tonPowerSupplyOn.Q
THEN
	udnErrorNo := 2; 								(* Set error number *)
	sErrorMsg := 'Power supply error';
END_IF
(*
IF lrSetTemp > 0
     AND lrActTemp > lrMaxTemp
THEN
	udnErrorNo := 2; 								(* Set error number *)
	sErrorMsg := 'Temperatur over range';
END_IF
*)

bError := udnErrorNo <> 0;

fbReadyDelay(
	bEnable := TRUE,
	bIn := bPowerOn,
	tDelay := tReadyDelay
);

IF lrSetTemp <> 0
     AND bAutoHand 			(* Automatic *)
THEN
	bReady := bPowerOn
			   AND lrActTemp >= lrSetTemp;
ELSE
	bReady := fbReadyDelay.bOut;
END_IF

(* Scaling power *)
fbScalingSP(
	bEnable := TRUE,
	lrInput := lrSPPower, (* [%] *)
	lrXLowLimit := 0, (* [%] *)
	lrXUpperLimit := 100, (* [%] *)
	lrYLowLimit := lrPowerMin, (* 16#0000 = 0 [V] *)
	lrYUpperLimit := lrPowerMax, (* 16#7FFF = 10 [V] *)
	usiPrecision := 2
);
unCVPower := LREAL_TO_UINT(fbScalingSP.lrOutputPV);

END_FUNCTION_BLOCK

// ---- POUs/Tc2 Objects/Automation/Force/FB_ForceReg.TcPOU
FUNCTION_BLOCK FB_ForceReg
VAR_INPUT
	rVelocityMax			:REAL := 10.0;
	rVelocityMin			:REAL := 0.0;
	PID_Reg: FB_PID_Regler;
	SollForceInt: INT := 20;
	IstForceInt: INT := 20;
	bRegelung: BOOL := FALSE;
	PWM_Aus: INT := 0;
	Force_Aus: REAL := 0.0;
	Simulation: BOOL := FALSE;
END_VAR
VAR_OUTPUT
	ForceOK: BOOL := FALSE;
	ForceOn: BOOL := FALSE;
	ForceLeistung: REAL := 0.0;
END_VAR
VAR
	PWM_Inc: INT := 0;
	PWM_Max: INT := 200;
	ForceModellReal: REAL := 0.0;
	K_Modell: REAL := 0.1;
	K_Modell_EM: REAL := 0.9;
	Force_Normal: REAL := 19.0;
	ForceModellInt: INT := 0;
	T_Modell: REAL := 360.0;
	bfirstCycle: BOOL := TRUE;
END_VAR

IF bFirstCycle THEN 				 (* Anfangsinitialisierungen *)

	PWM_Inc := 0;

	PID_Reg	(	
		fMax:=INT_TO_REAL(PWM_Max) ,
		fMin := 0.0,
		fD_Max := 1.0E10,
		fD_Min := -1.0E10,
		fKr := 1.0,
		fTN := 0.0,
		fTv := 0.0,
		fTau := 0.0,
		fOff := 0.0,
		fTab := 2.0,
		fState :=0.0,
		fIntegral := 0.0,
		fSoll := 0.0,
		fIst := 0.0
	);

	K_Modell 		:= EXP(-0.01/T_Modell);
	K_Modell_EM 	:= 1.0 - K_Modell;
	
	bFirstCycle:=FALSE;
END_IF

(* Zähler füR PID 0 incrementieren *)
PWM_Inc := 	PWM_Inc  + 1;

(* Regelung für PID 0 aufrufen *)
IF (PWM_Inc >= PWM_Max ) 
THEN
	PWM_Inc :=  0;

	(* Hier Regler einbauen *)
	IF bRegelung 
	THEN
		IF Simulation 
		THEN
			PID_Reg(fSoll:=SollForceInt, fIst:=ForceModellInt);
		ELSE
			PID_Reg(fSoll:=SollForceInt, fIst:=IstForceInt);
		END_IF
	
		PWM_Aus :=  REAL_TO_INT(PID_Reg.fAus);
		Force_Aus :=  PID_Reg.fAus;
		ForceOK := PID_Reg.bRegOK;
	ELSE
		PID_Reg.fIntegral := 0.0;
		PID_Reg(fSoll:=0.0, fIst:=0.0);
		PWM_Aus :=  0;
		Force_Aus :=  0.0;
		ForceOK := TRUE;
	
	END_IF

	IF ( PWM_Aus > PWM_Max ) THEN PWM_Aus:= PWM_Max; END_IF
	IF ( PWM_Aus < 0      ) THEN PWM_Aus := 0; END_IF

	IF ( Force_Aus > rVelocityMax ) THEN Force_Aus := rVelocityMax; END_IF
	IF ( Force_Aus < rVelocityMin ) THEN Force_Aus := rVelocityMin; END_IF

END_IF

(* PWM für PID  ausgeben == Inaktivierungsstrecke*)

ForceOn := FALSE;
IF (  PWM_Aus > PWM_Inc ) 
THEN		
	ForceOn := TRUE;        
END_IF

IF Simulation
THEN
	ForceModellReal := K_Modell*ForceModellReal;
	IF (  PWM_Aus > PWM_Inc ) THEN		ForceModellReal := K_Modell_EM*ForceModellReal;       END_IF
	ForceModellReal  := ForceModellReal + Force_Normal;
	ForceModellInt	:=REAL_TO_INT(ForceModellReal*10.0);
END_IF

END_FUNCTION_BLOCK

// ---- POUs/Tc2 Objects/Automation/Force/FB_PID_Regler.TcPOU
FUNCTION_BLOCK FB_PID_Regler
VAR_INPUT
	fSoll: REAL;
	fIst: REAL;
	fMax: REAL := 1.0;
	fMin: REAL := 0.0;
	fD_Max: REAL := 1.0;
	fD_Min: REAL := 0.0;
	fKr: REAL;
	fTn: REAL;
	fTv: REAL;
	fTau: REAL;
	fOff: REAL;
	fTab: REAL;
	fState: REAL;
	fIntegral: REAL;
END_VAR
VAR_OUTPUT
	bRegOK: BOOL := FALSE;
	fAus: REAL;
END_VAR
VAR
	fU: REAL;
	fU_Max: REAL;
	fU_Min: REAL;
	fU_Pd: ARRAY[1..2] OF REAL;
	fU_I: ARRAY[1..2] OF REAL;
	fE: ARRAY[1..4] OF REAL;
	fP: ARRAY[1..2] OF REAL;
	fQ: ARRAY[1..6] OF REAL;
	cMax: REAL;
	cMin: REAL;
	cD_Max: REAL := 1.0;
	cD_Min: REAL := 0.0;
	cKr: REAL;
	cTn: REAL;
	cTv: REAL;
	cTau: REAL;
	cOff: REAL;
	cTab: REAL;
	cState: REAL;
	cIntegral: REAL;
	nReg_Typ: INT;
	RegMaxAbweichung: REAL := 20.0;
END_VAR
VAR CONSTANT
	D_REG_I :INT:= 0;
	D_REG_M :INT := 1;
	D_REG_V :INT := 2;
	D_REG :INT := 4;
	I_REG :INT:= 8;
	P_REG :INT := 16;
	PD_I_REG :INT := 20;
	PD_M_REG :INT := 21;
	PD_V_REG :INT := 22;
	PI_REG :INT := 24;
	PID_I_REG :INT := 28;
	PID_M_REG :INT := 29;
	PID_V_REG :INT := 30;
	SET_MIN_MAX :INT := 101;
	ReglerResetState :INT := 102;
	ReglerInit :INT := 103;
	ReglerSet :INT := 104;
	ReglerCalculate :INT := 105;
END_VAR


IF (cMax  <>  fMax) 	THEN cMax := fMax; 	END_IF		 (*  Maximum                            *)
IF (cMin  <>  fMin) 	THEN cMin := fMin; 	END_IF	 	 (*  Minimum                            *)
IF (cD_Max  <>  fD_Max) 	THEN cD_Max := fD_Max; 	END_IF	 	 (*  Maximum der Änderung               *)
IF (cD_Min  <>  fD_Min) 		THEN cD_Min := fD_Min; 	END_IF	 	  (*  Minimum der Änderung               *)

IF ( (cState <>  fState) OR (cIntegral <>  fIntegral)) 		THEN
	cState := fState;
	cIntegral := fIntegral;
	fU := cState;
	fU_I[1] := fU_I[2] := cIntegral;
	fU_Pd[2] := fU_Pd[1] := 0.0;
	fE[4]		:=	fE[3]	:=	fE[2]		:=	fE[1]		:= 	0.0;
END_IF	 	  (*   Änderung Integral      *)

IF (  (cKr  <>  fKr) OR (cTn <> fTn) OR (cTv <> fTv) OR (cTau <> fTau)  OR (cOff <> fOff) OR (cTab <> fTab) ) THEN

     		cKr  := fKr;      (*  Verstärkung                       *)
		cTn  := fTn;      (*  Nachstellzeit                     *)
    		cTv  := fTv;      (*  Vorstellzeit                      *)
    		cTau := fTau;    (*  Tau                               *)
    		cOff := fOff;     (*  Offset                            *)

    		cTab := fTab;

(*    ReglerResetState(0.0, 0.0, p_r);           (*** Rücksetzen der Reglergrößen ***) *)
                  IF ( cTn = 0.0 ) THEN 	fU := fU_I[1] := fU_I[2] := 	fU_Pd[2] := fU_Pd[1] := 	fE[4]		:=	fE[3]	:=	fE[2]		:=	fE[1]		:= 	0.0;  END_IF

    		fP[1] := fP[2] := 0;         (*** Rücksetzen der Parameter ***)
    		fQ[1] := fQ[2] := fQ[3] := fQ[4] := fQ[5] := fQ[6] := 0;

    		nReg_Typ := 0;
    		IF ( cKr > 0 ) THEN nReg_Typ := nReg_Typ + P_REG;   END_IF  (*** Ermittlung der Reglertyps***)
    		IF ( cTn > 0 ) THEN nReg_Typ := nReg_Typ +  I_REG; END_IF
    		IF ( cTv > 0 ) THEN
      			 nReg_Typ := nReg_Typ + D_REG;
       			IF (cTau = 0) THEN nReg_Typ := nReg_Typ + D_REG_I;  END_IF(*** Ideale Differenz ***)
       			IF (cTau <  0) THEN nReg_Typ := nReg_Typ + D_REG_M;  END_IF(*** Gemittelte Differenz ***)
       			IF (cTau >  0) THEN nReg_Typ := nReg_Typ + D_REG_V;  END_IF(*** Verzögerte Differenz ***)
    		END_IF

		CASE nReg_Typ OF                  (*** Berechnung der Parameter ***)
		    P_REG :        (*** P-Regler ***********************************)
		       fQ[1] := cKr;
		    PI_REG :       (*** PI-Regler **********************************)
		       fQ[1] := cKr;

		       fQ[6] := cKr*cTab/cTn;
		    PD_I_REG :     (*** PD-Regler,      ideale Differenz  **********)
		       fQ[1] :=  cKr*cTv/cTab + cKr;
		       fQ[2] := -cKr*cTv/cTab;
		    PD_M_REG :     (*** PD-Regler,  gemittelte Differenz  **********)
		       fQ[1] :=  cKr*(1.0+cTv/6.0/cTab);
		       fQ[2] :=  cKr*cTv/2.0/cTab;
		       fQ[3] := -fQ[2];
		       fQ[4] :=  fQ[3]/3;
		    PD_V_REG :     (*** PD-Regler,  verzögerte Differenz  **********)
		       fP[1] := EXP(-cTab/cTau);

		       fQ[1] :=   cKr + cKr*cTv/cTau;
		       fQ[2] :=  -cKr - cKr*cTv/cTau + cKr*(1.0 - fP[1]) ;
		    PID_I_REG :    (*** PID-Regler,     ideale Differenz  **********)
		       fQ[1] :=  cKr*cTv/cTab + cKr;
		       fQ[2] := -cKr*cTv/cTab;

		       fQ[6] :=  cKr*cTab/cTn;
		    PID_M_REG :    (*** PID-Regler, gemittelte Differenz  **********)
		       fQ[1] :=  cKr*cTv/6/cTab + cKr;
		       fQ[2] :=  cKr*cTv/2/cTab;
		       fQ[3] := -fQ[2];
		       fQ[4] :=  fQ[3]/3;

		       fQ[6] :=  cKr*cTab/cTn;
		    PID_V_REG :    (*** PID-Regler, verzögerte Differenz  **********)
		       fP[1] :=  EXP(-cTab/cTau);

		       fQ[1] :=   cKr + cKr*cTv/cTau;
		       fQ[2] :=  -cKr - cKr*cTv/cTau + cKr*(1.0 - fP[1]) ;

		       fQ[6] :=  cKr*cTab/cTn;
		    I_REG :        (*** I-Regler ***********************************)
		       fQ[6] :=  cTab/cTn;

		END_CASE
END_IF


	fE[1] := fSoll - fIst;       	   (*** Regelabweichung ***)
	IF ( ABS(fE[1]) < RegMaxAbweichung ) THEN bRegOK := TRUE; ELSE bRegOK := FALSE; END_IF

	fU_Max := fU + cD_Max;   (*** dynamische Stellbegrenzung ***)
	IF (fU_Max > cMax) THEN fU_Max := cMax; END_IF

    	fU_Min := fU + cD_Min;
	IF (fU_Min < cMIN) THEN fU_Min := cMIN; END_IF
			                                          (*** Reglergleichung füR P- und D-Anteil***)
    	fU := fU_Pd[1] := fP[1]*fU_Pd[2] +   fQ[1]*fE[1] + fQ[2]*fE[2] +  fQ[3]*fE[3] + fQ[4]*fE[4];

                                          (*** Reglergleichung mit altem I-Anteil***)
    	fU := fU + fU_I[2];
                                      (*** Begrenzung der Stellgröße ***)
    	IF ( fU  > (fU_Max - cOff) ) THEN
             fU := fU_Max - cOff;
	ELSE
         		IF ( fU < (fU_Min - cOff) ) THEN
                		fU := fU_Min - cOff;
	         ELSE
                                          (*** Reglergleichung für I-Anteil***)
			fU_I[1] := fU_I[2] + fQ[6]*fE[1];
                                          (*** Gesamt-Reglergleichung ***)
			fU := (fU_Pd[1] + fU_I[1]);

                                      (*** Begrenzung der Stellgröße ***)
			IF ( fU > (fU_Max - cOff) ) THEN
                   		fU := fU_Max - cOff;
	                   	fU_I[1]  := fU - fU_Pd[1];
			ELSE
         		          	IF ( fU < (fU_Min - cOff) ) THEN
                   			fU := fU_Min - cOff;
		         		         fU_I[1]  := fU - fU_Pd[1];
	         		      	END_IF
         		   	END_IF
         		END_IF
    	END_IF                                          (*** Umspeichern der Regelgrößen ***)
	fU_Pd[2] := fU_Pd[1];
	fU_I[2]  := fU_i[1];

	fE[4] := fE[3];
	fE[3] := fE[2];
	fE[2] := fE[1];

                                        (*** Übergabe der Stellgröße ***)
	fAus := fU + cOff;

END_FUNCTION_BLOCK

// ---- POUs/Tc2 Objects/Automation/Force/FB_FORCE_REF.TcPOU
FUNCTION_BLOCK FB_FORCE_REF
VAR_INPUT
	unForceMeasureType			:UINT;								(* Type of force measure system. 1: Simple mA,  2: EL3351 3: EL3356 *)

	fbForceSimple				:FB_ScalingOffset;

	lrForceMin					:LREAL;								(* Force min [mA] 16#0000 = 4 [mA] *)
	lrForceMax	 				:LREAL;								(* Force max [mA] 16#7FFF = 20 [mA] *)
	lrForceMinN					:LREAL;								(* Force min [N] *)
	lrManualForceMaxN			:LREAL;								(* Force max [N] *)
	lrAutoForceMaxN				:LREAL;								(* Force max [N] *)

	fbForceEL3356				:FB_EL3356;

	stRefSettingsEL3356			:ST_EL3356CoeInfo;					(* Reference settings of EL3356 force input modul *)
	stActSettingsEL3356			:ST_EL3356CoeInfo;					(* Actual settings of EL3356 force input modul *)

	stTerminalStateEL3356			AT %I*:ST_TerminalState;				(* Terminal state EL3356 *)
	stChannelStateEL3356			AT %I*:ST_EL3356ChannelState;		(* Channel state EL3356 *)
	stChannelCtrlEL3356			AT %Q*:ST_EL3356ChannelCtrl;			(* Channel control EL3356 *)

	stForceToPlc					AT %I*:ST_FORCETOPLC;
	stPlcToForce					AT %Q*:ST_PLCTOFORCE;
END_VAR
VAR_OUTPUT

END_VAR
VAR_IN_OUT

END_VAR
VAR

END_VAR

;

END_FUNCTION_BLOCK

// ---- POUs/Tc2 Objects/Automation/Heater/FB_Heater.TcPOU
FUNCTION_BLOCK FB_Heater
(*

The function block used to control heater.

Constructor: 		Patryk Panylo
Company:		E. Riexinger GmbH
Date:			07.09.2018
Version:			1.00

Date:			Revision:		Who:				Comment
xx.xx.xxxx			1.01									

*)
VAR_INPUT
	(* Input variables / Eingang Variablen *)
	bEnable							:BOOL;						(* Function block enable *)
	bNoEStop						:BOOL;						(* No ermergency Stop / Keine Notaus *)
	bPowerSupplyOn					:BOOL;						(* Power supply on / Leitung eingeschaltet *)
	bLightCurtainOK					:BOOL;						(* Light curtain ok / Freigabe Lichtschranke i.o *)
	bReset							:BOOL;						(* Controller reset *)
	bAutoHand						:BOOL;						(* Auto := TRUE, Hand := FALSE *)
	bHandOn						:BOOL;						(* Heater on/off in manual mode with rising edge *)
	bAutoOn							:BOOL;						(* Heater on/off in auto mode rising edge *)
	bAutoOff							:BOOL;						(* Heater off in auto mode with rising edge *)
	bReleaseOn						:BOOL;						(* Release on *)
	bCtrlInterrupt						:BOOL;						(* Control interrupt *)
	lrSPPower						:LREAL;						(* Setpoint of power 0 - 100 % *)
	bEnAutoCtrlOff					:BOOL := FALSE;				(* Auto off enable*)
	tCtrlPowerOff						:TIME := t#90s;				(* Time to switch controller power off *)
	tCtrlPowerOn						:TIME := t#90s;				(* Time to switch controller power on *)
	lrPowerMin						:LREAL;						(* Power minimum *)
	lrPowerMax						:LREAL;						(* Power maximum *)
	lrSetTemp						:LREAL;						(* Set temperature *)
	lrActTemp						:LREAL;						(* Actual temperature *)
	lrMaxTemp						:LREAL;						(* Maximal temperature *)
	tReadyDelay						:TIME := T#5s;				(* Ready delay*)
	tTimeOut							:TIME := T#5s;				(* TimeOut *)
END_VAR
VAR_OUTPUT
	(* Output variables / Ausgang Variablen *)
	bPowerOn						:BOOL;						(* Power on *)
	unCVPower						:UINT;						(* Current value of power 0 - 10 V *)
	bReady 							:BOOL;						(* Heater ready *)
	bError							:BOOL;						(* Program error  *)
	udnErrorNo						:UDINT;						(* Error number *)
	sErrorMsg						:STRING; 					(* Error message *)
END_VAR
VAR_IN_OUT
	(* Input Output variables / Ausgang Variablen *)

END_VAR
VAR
	(* Enummerations *)

	(* Variables *)
	bReleasePowerOn				:BOOL;

	bFirstTime						:BOOL;

	(* References *)

	(* Interfaces *)

	(* Instances *)
	tonWatchDog						:TON;
	tonPowerSupplyOn				:TON;
	fbCtrlPowerOff					:FB_SignalHandlingDelay;
	fbCtrlPowerOn					:FB_SignalHandlingDelay;
	fbScalingSP						:FB_Scaling;
	fbReadyDelay					:FB_SignalHandlingDelay;

	rtHandOn						:R_TRIG;
	rtAutoOn							:R_TRIG;
	rtAutoOff							:R_TRIG;
END_VAR
VAR CONSTANT

END_VAR


IF NOT bEnable
THEN
	bPowerOn := FALSE;				(* Power on *)
 	unCVPower := 0;					(* Current value of power 0 - 100 % *)
	bReady := TRUE;				(* Heater enabled *)
	bError := FALSE;					(* Program error  *)
	udnErrorNo := 0;					(* Error number *)
	sErrorMsg := ''; 					(* Error message *)
	tonWatchDog(IN := FALSE);

	bFirstTime := FALSE;
	RETURN;
END_IF

IF NOT bFirstTime
THEN
	bReleasePowerOn := TRUE;

	bPowerOn := FALSE;				(* Powr on *)
 	unCVPower := 0;					(* Current value of power 0 - 100 % *)
	bReady := FALSE;				(* Heater enabled *)

	bFirstTime := TRUE;
END_IF

(* Controller automatic off *)
fbCtrlPowerOff(
	bEnable := TRUE,
	bIn := bEnAutoCtrlOff
		  AND bPowerOn,
	tDelay := tCtrlPowerOff
);

fbCtrlPowerOn(
	bEnable := TRUE,
	bIn := NOT bPowerOn					(* Ctrl disabled *)
		  AND NOT bReleasePowerOn,
	tDelay := tCtrlPowerOn
);

IF NOT bNoEStop
     OR NOT bPowerSupplyOn
     OR NOT bLightCurtainOK
     OR bError
     OR bCtrlInterrupt
     OR fbCtrlPowerOff.bOut
THEN
	bReleasePowerOn := FALSE;
	bPowerOn := FALSE;

ELSIF fbCtrlPowerOn.bOut
THEN
	bReleasePowerOn := TRUE;
END_IF

